(* IEC 61131-3 sources: daoli-st-library/DL_Process (part 9) *)

(* ---- FC_DL_AnodizeBathChargeCalc.st ---- *)
(*
  Component : FC_DL_AnodizeBathChargeCalc
  Category  : DL_Process
  Type      : FC
  Complexity: C2
  VERSION   : v1.0.0
  功能      : 阳极氧化槽法拉第电量核算：Q = I·t，换算电量密度与膜厚，并按电流效率由目标膜厚反算所需时间。
  开源溯源  : 道莅原创 clean-room 自研（无外部代码引用）｜License: MIT
  边界条件  : ① 氧化面积、电流效率、单位电量膜厚系数须 > 1e-9 且效率不超过 100 %，否则返回哨兵 -1；
              ② 电流为 0 时膜厚为 0 且反算时间回 0（合法空工况，xValid 置真）；
              ③ 反算时间不下发负值，目标膜厚 <= 0 时直接回 0。
*)
FUNCTION FC_DL_AnodizeBathChargeCalc : REAL
VAR_INPUT
    fCurrentA     : REAL;   (* 整流器输出电流 [A] Rectifier output current *)
    fAreaDm2      : REAL;   (* 氧化有效面积 [dm²] Effective anodizing area *)
    fTimeS        : REAL;   (* 通电时长 [s] Energizing time *)
    fEffPct       : REAL;   (* 电流效率 [%] Current efficiency *)
    fUmPerAsDm2   : REAL;   (* 单位电量膜厚系数 [μm/(A·s/dm²)] Film thickness per charge density *)
    fThickTargetUm: REAL;   (* 目标膜厚 [μm] Target film thickness *)
END_VAR
VAR_OUTPUT
    fChargeC       : REAL;  (* 累计电量 [C] Accumulated charge *)
    fChgDensAsDm2  : REAL;  (* 电量密度 [A·s/dm²] Charge density *)
    fFilmUm        : REAL;  (* 实测对应膜厚 [μm] Film thickness from charge *)
    fTimeForTargetS: REAL;  (* 达目标膜厚所需时间 [s] Time to reach target thickness *)
    xValid         : BOOL;  (* 计算有效性标志 [-] Calculation valid flag *)
END_VAR
VAR CONSTANT
    DL_EPS      : REAL := 1.0E-9;   (* 除零判定容差 [无量纲] Divide-by-zero tolerance *)
    DL_PCT_BASE : REAL := 100.0;    (* 百分比基准 [%] Percent base *)
    DL_ZERO     : REAL := 0.0;      (* 零常量 [无量纲] Zero constant *)
END_VAR
VAR
    fDensADm2 : REAL;   (* 电流密度 [A/dm²] Current density *)
    fEffUnit  : REAL;   (* 效率折算系数 [-] Efficiency as fraction *)
END_VAR
(* 出口预置：五出口统一预置 *)
fChargeC := 0.0; fChgDensAsDm2 := 0.0; fFilmUm := 0.0; fTimeForTargetS := 0.0; xValid := FALSE;
(* 非有限拦截：自反判 NaN，自身差值判 Inf *)
IF (fCurrentA <> fCurrentA) OR ((fCurrentA - fCurrentA) <> 0.0)
   OR (fAreaDm2 <> fAreaDm2) OR ((fAreaDm2 - fAreaDm2) <> 0.0)
   OR (fTimeS <> fTimeS) OR ((fTimeS - fTimeS) <> 0.0)
   OR (fEffPct <> fEffPct) OR ((fEffPct - fEffPct) <> 0.0)
   OR (fUmPerAsDm2 <> fUmPerAsDm2) OR ((fUmPerAsDm2 - fUmPerAsDm2) <> 0.0) THEN
    FC_DL_AnodizeBathChargeCalc := -1.0;  (* 哨兵 -1：输入非有限 / Sentinel -1 non-finite *)
    RETURN;
END_IF
(* 组态域闸：面积与系数为除子/比例基，电流与时长须非负，效率须在 (0,100] *)
IF (fAreaDm2 <= DL_EPS) OR (fUmPerAsDm2 <= DL_EPS) OR (fEffPct <= DL_ZERO)
   OR (fEffPct > DL_PCT_BASE) OR (fCurrentA < DL_ZERO) OR (fTimeS < DL_ZERO) THEN
    FC_DL_AnodizeBathChargeCalc := -1.0;  (* 哨兵 -1：组态非法 / Sentinel -1 bad config *)
    RETURN;
END_IF
fEffUnit := fEffPct / DL_PCT_BASE;             (* 效率折算 [-] / Efficiency as fraction *)
(* 电量：Q = I·t [C] = [A·s] *)
fChargeC := fCurrentA * fTimeS;
(* 电量密度与电流密度：分母面积已过域闸 *)
fChgDensAsDm2 := fChargeC / fAreaDm2;
fDensADm2 := fCurrentA / fAreaDm2;
(* 膜厚：δ = 电量密度 × 单位膜厚系数 × 电流效率 [μm] *)
fFilmUm := fChgDensAsDm2 * fUmPerAsDm2 * fEffUnit;
(* 反算时间：t = 目标膜厚 / (电流密度 × 系数 × 效率)，电流密度为 0 时回 0 *)
IF (fDensADm2 > DL_EPS) AND (fThickTargetUm > DL_ZERO) THEN
    fTimeForTargetS := fThickTargetUm / (fDensADm2 * fUmPerAsDm2 * fEffUnit);
END_IF
xValid := TRUE;                                (* 链路有效 / Chain valid *)
FC_DL_AnodizeBathChargeCalc := fFilmUm;        (* 返回膜厚 [μm] / Return film thickness *)
END_FUNCTION

(* ---- FC_DL_AnodizeSealBoilTimeCalc.st ---- *)
(*
  Component : FC_DL_AnodizeSealBoilTimeCalc
  Category  : DL_Process
  Type      : FC
  Complexity: C1
  VERSION   : v1.0.0
  功能      : 沸水封孔时间核算：按膜厚乘单位膜厚基准时间，再叠加温度窗口修正，判定 pH/温度窗口与最终封孔合格性。
  开源溯源  : 道莅原创 clean-room 自研（无外部代码引用）｜License: MIT
  边界条件  : ① 膜厚与单位膜厚时间须 > 1e-9，否则返回哨兵 -1；
              ② pH 窗口 5.5~6.5、温度窗口 95~100 °C，任一越窗即判不合格但不拒算；
              ③ 温度修正系数钳位 1.0~2.0，温度偏低延长封孔时间。
*)
FUNCTION FC_DL_AnodizeSealBoilTimeCalc : REAL
VAR_INPUT
    fFilmUm    : REAL;   (* 氧化膜厚 [μm] Oxide film thickness *)
    fBathTempC : REAL;   (* 封孔槽液温度 [°C] Sealing bath temperature *)
    fPh        : REAL;   (* 封孔槽液 pH [-] Sealing bath pH *)
    fMinPerUm  : REAL;   (* 单位膜厚基准封孔时间 [min/μm] Base sealing time per um *)
    fFilmMinUm : REAL;   (* 可封孔最小膜厚 [μm] Minimum sealable film thickness *)
END_VAR
VAR_OUTPUT
    fSealTimeMin : REAL;  (* 封孔时间 [min] Sealing time *)
    fTempCoef    : REAL;  (* 温度修正系数 [-] Temperature correction coefficient *)
    xWindowOk    : BOOL;  (* pH 与温度窗口合格标志 [-] Window valid flag *)
    xQualified   : BOOL;  (* 封孔合格标志 [-] Sealing qualified flag *)
    xValid       : BOOL;  (* 计算有效性标志 [-] Calculation valid flag *)
END_VAR
VAR CONSTANT
    DL_EPS      : REAL := 1.0E-9;   (* 除零判定容差 [无量纲] Divide-by-zero tolerance *)
    DL_PH_LO    : REAL := 5.5;      (* pH 窗口下限 [-] pH window lower bound *)
    DL_PH_HI    : REAL := 6.5;      (* pH 窗口上限 [-] pH window upper bound *)
    DL_TMP_LO   : REAL := 95.0;     (* 温度窗口下限 [°C] Temperature window lower bound *)
    DL_TMP_HI   : REAL := 100.0;    (* 温度窗口上限 [°C] Temperature window upper bound *)
    DL_TMP_REF  : REAL := 100.0;    (* 温度修正基准 [°C] Temperature reference *)
    DL_TMP_SLOPE: REAL := 0.25;     (* 每 10 °C 温度修正量 [-] Slope per 10 degC *)
    DL_COEF_MAX : REAL := 2.0;      (* 温度修正上限 [-] Temperature coefficient clamp *)
END_VAR
VAR
    fGapC : REAL;   (* 相对基准温度的温差 [°C] Temperature gap from reference *)
END_VAR
(* 出口预置：五出口统一预置 *)
fSealTimeMin := 0.0; fTempCoef := 1.0; xWindowOk := FALSE; xQualified := FALSE; xValid := FALSE;
(* 非有限拦截：自反判 NaN，自身差值判 Inf *)
IF (fFilmUm <> fFilmUm) OR ((fFilmUm - fFilmUm) <> 0.0)
   OR (fBathTempC <> fBathTempC) OR ((fBathTempC - fBathTempC) <> 0.0)
   OR (fPh <> fPh) OR ((fPh - fPh) <> 0.0) THEN
    FC_DL_AnodizeSealBoilTimeCalc := -1.0;  (* 哨兵 -1：输入非有限 / Sentinel -1 non-finite *)
    RETURN;
END_IF
(* 组态域闸：膜厚与单位膜厚时间均为比例基 *)
IF (fFilmUm < DL_EPS) OR (fMinPerUm <= DL_EPS) THEN
    FC_DL_AnodizeSealBoilTimeCalc := -1.0;  (* 哨兵 -1：组态非法 / Sentinel -1 bad config *)
    RETURN;
END_IF
(* 窗口判定：pH 与温度双窗口，任一越窗即判不合格（不拒算，便于上位诊断） *)
IF (fPh >= DL_PH_LO) AND (fPh <= DL_PH_HI)
   AND (fBathTempC >= DL_TMP_LO) AND (fBathTempC <= DL_TMP_HI) THEN
    xWindowOk := TRUE;
END_IF
(* 温度修正：低于基准温度每 10 °C 延长 25 %，双侧钳位 *)
fGapC := DL_TMP_REF - fBathTempC;
IF fGapC > 0.0 THEN
    fTempCoef := 1.0 + (fGapC / 10.0) * DL_TMP_SLOPE;
ELSE
    fTempCoef := 1.0;                       (* 达到或高于基准：不缩短，防欠封 *)
END_IF
IF fTempCoef > DL_COEF_MAX THEN
    fTempCoef := DL_COEF_MAX;               (* 上限钳位 [-] / Upper clamp *)
END_IF
(* 封孔时间：t = 膜厚 × 单位膜厚时间 × 温度修正，分母均已过域闸 *)
fSealTimeMin := fFilmUm * fMinPerUm * fTempCoef;
(* 合格判定：窗口合格且膜厚达可封孔最小值 *)
xQualified := xWindowOk AND (fFilmUm >= fFilmMinUm);
xValid := TRUE;                             (* 链路有效 / Chain valid *)
FC_DL_AnodizeSealBoilTimeCalc := fSealTimeMin;  (* 返回封孔时间 [min] / Return sealing minutes *)
END_FUNCTION

(* ---- FC_DL_AustenitizeHoldTimeCalc.st ---- *)
(*
  Component : FC_DL_AustenitizeHoldTimeCalc
  Category  : DL_Process
  Type      : FC
  Complexity: C2
  VERSION   : v1.0.0
  功能      : 奥氏体化保温时间核算：按有效厚度乘以单位厚度基准时间，再叠加厚度分段系数、升温速率修正与目标温度修正。
  开源溯源  : 道莅原创 clean-room 自研（无外部代码引用）｜License: MIT
  边界条件  : ① 有效厚度/升温速率/单位厚度时间均须 > 1e-9，否则返回哨兵 -1；
              ② 厚度分三段（<=25 / <=50 / >50 mm），系数逐段离散，段内不插值；
              ③ 升温速率修正与温度修正均双侧钳位，防经验式外推发散。
*)
FUNCTION FC_DL_AustenitizeHoldTimeCalc : REAL
VAR_INPUT
    fThkMm      : REAL;   (* 工件有效厚度 [mm] Effective thickness *)
    fRateCmin   : REAL;   (* 实际升温速率 [°C/min] Actual heating rate *)
    fRateRefCmin: REAL;   (* 参考升温速率（分段基准） [°C/min] Reference heating rate *)
    fTargetC    : REAL;   (* 目标奥氏体化温度 [°C] Target austenitizing temperature *)
    fTempRefC   : REAL;   (* 参考目标温度（分段基准） [°C] Reference target temperature *)
    fMinPerMm   : REAL;   (* 单位厚度基准保温时间 [min/mm] Base hold time per mm *)
END_VAR
VAR_OUTPUT
    fHoldMin   : REAL;    (* 保温时间计算结果 [min] Computed hold time *)
    fThkCoef   : REAL;    (* 厚度分段系数 [-] Thickness segment coefficient *)
    fRateCoef  : REAL;    (* 升温速率修正系数 [-] Heating rate correction coefficient *)
    xValid     : BOOL;    (* 计算有效性标志 [-] Calculation valid flag *)
END_VAR
VAR CONSTANT
    DL_EPS       : REAL := 1.0E-9;   (* 除零判定容差 [无量纲] Divide-by-zero tolerance *)
    DL_RATE_MIN  : REAL := 0.80;     (* 速率修正下限 [-] Rate correction lower clamp *)
    DL_RATE_MAX  : REAL := 1.30;     (* 速率修正上限 [-] Rate correction upper clamp *)
    DL_TEMP_K    : REAL := 0.002;    (* 目标温度每 °C 修正斜率 [1/°C] Temperature slope *)
    DL_THK_MID   : REAL := 25.0;     (* 厚度分段第一界 [mm] First thickness boundary *)
    DL_THK_HIGH  : REAL := 50.0;     (* 厚度分段第二界 [mm] Second thickness boundary *)
END_VAR
(* 出口预置：全出口统一预置 *)
fHoldMin := 0.0; fThkCoef := 1.0; fRateCoef := 1.0; xValid := FALSE;
(* 非有限拦截：自反判 NaN，自身差值判 Inf *)
IF (fThkMm <> fThkMm) OR ((fThkMm - fThkMm) <> 0.0)
   OR (fRateCmin <> fRateCmin) OR ((fRateCmin - fRateCmin) <> 0.0)
   OR (fRateRefCmin <> fRateRefCmin) OR ((fRateRefCmin - fRateRefCmin) <> 0.0)
   OR (fTargetC <> fTargetC) OR ((fTargetC - fTargetC) <> 0.0)
   OR (fTempRefC <> fTempRefC) OR ((fTempRefC - fTempRefC) <> 0.0)
   OR (fMinPerMm <> fMinPerMm) OR ((fMinPerMm - fMinPerMm) <> 0.0) THEN
    FC_DL_AustenitizeHoldTimeCalc := -1.0;  (* 哨兵 -1：输入非有限 / Sentinel -1 non-finite *)
    RETURN;
END_IF
(* 组态域闸：厚度、实际升温速率、单位厚度时间三者为除子或比例基 *)
IF (fThkMm <= DL_EPS) OR (fRateCmin <= DL_EPS) OR (fMinPerMm <= DL_EPS) THEN
    FC_DL_AustenitizeHoldTimeCalc := -1.0;  (* 哨兵 -1：组态非法 / Sentinel -1 bad config *)
    RETURN;
END_IF
(* 厚度分段系数：三段离散，段内不插值，防止经验式在厚壁区外推 *)
IF fThkMm <= DL_THK_MID THEN
    fThkCoef := 1.00;                       (* 薄件段 [-] / Thin section *)
ELSIF fThkMm <= DL_THK_HIGH THEN
    fThkCoef := 1.15;                       (* 中厚段 [-] / Medium section *)
ELSE
    fThkCoef := 1.35;                       (* 厚壁段（心部透热滞后） [-] / Thick section *)
END_IF
(* 升温速率修正：升温越慢，组织转变越充分，保温时间可缩短，双侧钳位 *)
fRateCoef := fRateRefCmin / fRateCmin;
IF fRateCoef < DL_RATE_MIN THEN
    fRateCoef := DL_RATE_MIN;               (* 下限钳位 [-] / Lower clamp *)
ELSIF fRateCoef > DL_RATE_MAX THEN
    fRateCoef := DL_RATE_MAX;               (* 上限钳位 [-] / Upper clamp *)
END_IF
(* 目标温度修正：温度偏低需延长保温 *)
IF fTargetC > fTempRefC THEN
    fHoldMin := fMinPerMm * fThkMm * fThkCoef * fRateCoef;
    fHoldMin := fHoldMin * (1.0 - (fTargetC - fTempRefC) * DL_TEMP_K);
ELSE
    fHoldMin := fMinPerMm * fThkMm * fThkCoef * fRateCoef;
    fHoldMin := fHoldMin * (1.0 + (fTempRefC - fTargetC) * DL_TEMP_K);
END_IF
(* 结果下钳位：保温时间不得为负，防温度修正项越界 *)
IF fHoldMin < DL_EPS THEN
    fHoldMin := DL_EPS;                     (* 非负钳位 [min] / Non-negative clamp *)
END_IF
xValid := TRUE;                             (* 链路有效 / Chain valid *)
FC_DL_AustenitizeHoldTimeCalc := fHoldMin;  (* 返回保温时间 [min] / Return hold minutes *)
END_FUNCTION

(* ---- FC_DL_BallMillPowerDrawCalc.st ---- *)
(*
  Name: FC_DL_BallMillPowerDrawCalc
  Category: DL_Process
  Version: 1.0.0
  Round: R89 / 2026-11-25
  开源溯源：clean-room 自研（族 矿山破碎筛分，ST 开源生态实测 0 命中，无外部代码引入）
  功能：球磨机轴功率与比能耗估算（筒径/筒长/转速率/装球率经验幂律），并折算单位给矿能耗。
  边界条件：① 五入参全部过非有限闸，任一非有限返回哨兵 -1；
            ② 筒径 0.5~8 m、筒长 0.5~15 m、临界转速率 30~100 %、装球率 10~55 % 为工程域，越域返回哨兵 -1；
            ③ 给矿量为 0 属正常运行工况（空转），比能耗输出 0 而不判非法，功率照常有效；
            ④ 幂次 2.5 以 D·D·SQRT(D) 展开实现，不引入 EXPT 原语（R140 委托纪律）。
  量纲自证：K[kW/m^3.5] × D^2.5[m^2.5] × L[m] = kW；转速率与装球率为无量纲百分比折算。
*)
FUNCTION FC_DL_BallMillPowerDrawCalc : REAL
VAR_INPUT
    fMillDiaM : REAL;        (* 磨机筒体有效内径 [m] Mill effective diameter [m] *)
    fMillLenM : REAL;        (* 磨机筒体有效长度 [m] Mill effective length [m] *)
    fSpeedPct : REAL;        (* 临界转速百分比 [%] Percent of critical speed [%] *)
    fMediaLoadPct : REAL;    (* 装球率（磨机容积占比） [%] Ball charge volume ratio [%] *)
    fFeedTph : REAL;         (* 给矿量 [t/h] Feed rate [t/h] *)
END_VAR
VAR_OUTPUT
    fPowerKW : REAL;         (* 磨机轴功率 [kW] Mill shaft power [kW] *)
    fSpecificKWhT : REAL;    (* 单位给矿能耗 [kWh/t] Specific energy per tonne [kWh/t] *)
    xValid : BOOL;           (* 计算有效性标志 [-] Calculation valid flag *)
END_VAR
VAR CONSTANT
    DL_EPS : REAL := 1.0E-9;        (* 除零判定容差 [-] Divide-by-zero tolerance *)
    DL_K_POWER : REAL := 26.0;      (* 功率经验系数 [kW/m^3.5] Empirical power coefficient *)
    DL_D_MIN : REAL := 0.5;         (* 筒径下限 [m] Diameter floor [m] *)
    DL_D_MAX : REAL := 8.0;         (* 筒径上限 [m] Diameter ceiling [m] *)
    DL_L_MIN : REAL := 0.5;         (* 筒长下限 [m] Length floor [m] *)
    DL_L_MAX : REAL := 15.0;        (* 筒长上限 [m] Length ceiling [m] *)
    DL_SPD_MIN : REAL := 30.0;      (* 转速率下限 [%] Speed ratio floor [%] *)
    DL_SPD_MAX : REAL := 100.0;     (* 转速率上限 [%] Speed ratio ceiling [%] *)
    DL_MED_MIN : REAL := 10.0;      (* 装球率下限 [%] Media load floor [%] *)
    DL_MED_MAX : REAL := 55.0;      (* 装球率上限 [%] Media load ceiling [%] *)
    DL_PCT : REAL := 100.0;         (* 百分数基准 [%] Percent base *)
END_VAR
VAR
    fD25 : REAL;    (* 筒径 2.5 次幂 [m^2.5] Diameter to the power 2.5 *)
    fKspd : REAL;   (* 转速率折算系数 [-] Speed ratio factor *)
    fKmed : REAL;   (* 装球率折算系数 [-] Media load factor *)
END_VAR
(* 出口预置：三出口统一预置（R256） *)
fPowerKW := 0.0; fSpecificKWhT := 0.0; xValid := FALSE;
(* 非有限闸：NaN 自反判 + Inf 差值自减判，五入参全枚举 *)
IF (fMillDiaM <> fMillDiaM) OR ((fMillDiaM - fMillDiaM) <> 0.0)
   OR (fMillLenM <> fMillLenM) OR ((fMillLenM - fMillLenM) <> 0.0)
   OR (fSpeedPct <> fSpeedPct) OR ((fSpeedPct - fSpeedPct) <> 0.0)
   OR (fMediaLoadPct <> fMediaLoadPct) OR ((fMediaLoadPct - fMediaLoadPct) <> 0.0)
   OR (fFeedTph <> fFeedTph) OR ((fFeedTph - fFeedTph) <> 0.0) THEN
    FC_DL_BallMillPowerDrawCalc := -1.0;    (* 哨兵 -1：入参非有限 / Sentinel -1, non-finite input *)
    RETURN;
END_IF
(* 组态域闸：几何与工艺参数逐项定域，给矿量允许为 0（空转） *)
IF (fMillDiaM < DL_D_MIN) OR (fMillDiaM > DL_D_MAX)
   OR (fMillLenM < DL_L_MIN) OR (fMillLenM > DL_L_MAX)
   OR (fSpeedPct < DL_SPD_MIN) OR (fSpeedPct > DL_SPD_MAX)
   OR (fMediaLoadPct < DL_MED_MIN) OR (fMediaLoadPct > DL_MED_MAX)
   OR (fFeedTph < 0.0) THEN
    FC_DL_BallMillPowerDrawCalc := -1.0;    (* 哨兵 -1：组态非法 / Sentinel -1, bad configuration *)
    RETURN;
END_IF
(* 幂次展开：D^2.5 = D·D·√D，量纲 m^2.5 *)
fD25 := fMillDiaM * fMillDiaM * SQRT(fMillDiaM);
(* 两百分比折算为无量纲系数 *)
fKspd := fSpeedPct / DL_PCT;
fKmed := fMediaLoadPct / DL_PCT;
(* 轴功率：K[kW/m^3.5] × D^2.5 × L × kspd × kmed，量纲收敛为 kW *)
fPowerKW := DL_K_POWER * fD25 * fMillLenM * fKspd * fKmed;
(* 比能耗：给矿为 0 时输出 0（除零保护，且空转不产比能耗事实） *)
IF fFeedTph > DL_EPS THEN
    fSpecificKWhT := fPowerKW / fFeedTph;   (* kW ÷ (t/h) = kWh/t *)
ELSE
    fSpecificKWhT := 0.0;                   (* 空转：无比能耗 / No specific energy at no feed *)
END_IF
xValid := TRUE;                             (* 链路有效 / Chain valid *)
FC_DL_BallMillPowerDrawCalc := fPowerKW;
END_FUNCTION

(* ---- FC_DL_BeamToppleRiskChk.st ---- *)
(*
  ============================================================
  组件名 : FC_DL_BeamToppleRiskChk
  分类   : DL_Process
  功能   : 横梁倾覆风险校核，按重心偏心放大力矩后折算横梁承载利用率并给出风险位
  复杂度 : C1
  版本   : 1.0.1
  作者   : 道莅工业代码库工厂 / R81
  日期   : 2026-11-24
  开源溯源 : clean-room（no upstream）—— 依据公开工程公式自研，未复制任何上游实现
  红线自检 : R1 无GVL/R2 无物理地址/R3 纯IEC/R4 防除零/R5 双语注释
  接口说明 :
      偏心系数 = 1 + |重心偏移|/横梁深度（v1.0.1 取绝对值：负偏移同样放大倾覆风险，
      修正原带符号实现导致负偏移时利用率被低估、风险漏报的缺陷），偏心为零时系数为 1。
      |重心偏移| > 梁深/2 视为不可信组态，直接置 bValid=FALSE 返回。
      有效载荷 = 载荷 * 偏心系数；利用率超过 85% 即判倾覆风险。
      利用率不做 100% 上限截断，超过 100% 的信息对诊断有价值，由调用侧自行显示。
  ============================================================
*)
FUNCTION FC_DL_BeamToppleRiskChk : BOOL
VAR_INPUT
    bEnable      : BOOL; // 使能：TRUE 时校核 / Enable: TRUE to check
    bErr         : BOOL; // 外部故障：TRUE 时立即退出并置结果无效 / External fault: TRUE aborts with invalid result
    rLoadKg      : REAL; // 实际载荷质量 [kg] / actual load mass [kg]
    rBeamCapKg   : REAL; // 横梁额定承载质量 [kg] / rated load capacity of the beam [kg]
    rCgOffset_mm : REAL; // 载荷重心相对横梁中心的偏移 [mm] / load centre of gravity offset from the beam centre [mm]
    rBeamDepth_mm : REAL; // 横梁截面深度 [mm] / beam section depth [mm]
END_VAR
VAR_OUTPUT
    rEccFactor : REAL; // 偏心放大系数 [无量纲] / eccentricity amplification factor [dimensionless]
    rEffLoadKg : REAL; // 折算有效载荷质量 [kg] / equivalent effective load mass [kg]
    rUtilPct   : REAL; // 承载利用率 [%] / utilisation of the rated capacity [percent]
    bRisk      : BOOL; // 倾覆风险：TRUE 表示利用率超过门限 / topple risk, TRUE when utilisation exceeds the limit
    bValid     : BOOL; // 输出有效：TRUE 表示结果可用 / Output valid
END_VAR
VAR CONSTANT
    DL_R_MAX    : REAL := 3.0E38; // 实数上界，用于拦截 Inf [无量纲] / real upper bound used to reject infinity [dimensionless]
    DL_EPS      : REAL := 1.0E-12; // 除零判定阈值 [无量纲] / division guard threshold [dimensionless]
    DL_RISK_PCT : REAL := 85.0;   // 倾覆风险门限 [%] / topple risk threshold [percent]
    DL_PCT      : REAL := 100.0;  // 百分数换算系数 [无量纲] / percentage scaling factor [dimensionless]
END_VAR
VAR
    _bFin : BOOL := FALSE; // 输入有限性判定结果 / input finiteness verdict
END_VAR

    // 段 1｜出口预置
    rEccFactor := 1.0;
    rEffLoadKg := 0.0;
    rUtilPct := 0.0;
    bRisk := FALSE;
    bValid := FALSE;
    // 段 2｜使能闸与外部故障闸
    IF NOT bEnable THEN
        RETURN;
    END_IF;
    IF bErr THEN
        RETURN;
    END_IF;
    // 段 3｜非有限闸
    _bFin := (rLoadKg = rLoadKg) AND (ABS(rLoadKg) <= DL_R_MAX) AND (rBeamCapKg = rBeamCapKg) AND (ABS(rBeamCapKg) <= DL_R_MAX) AND (rCgOffset_mm = rCgOffset_mm) AND (ABS(rCgOffset_mm) <= DL_R_MAX) AND (rBeamDepth_mm = rBeamDepth_mm) AND (ABS(rBeamDepth_mm) <= DL_R_MAX);
    IF NOT _bFin THEN
        RETURN;
    END_IF;
    // 段 4｜域闸：承载与横梁深度必须为正，载荷不得为负
    IF (ABS(rBeamCapKg) <= DL_EPS) OR (ABS(rBeamDepth_mm) <= DL_EPS) THEN
        RETURN;
    END_IF;
    IF (rBeamCapKg < 0.0) OR (rLoadKg < 0.0) OR (rBeamDepth_mm < 0.0) THEN
        RETURN;
    END_IF;
    // 段 4b｜偏心量域闸：|偏移| 超过梁深一半即视为不可信组态，直接置无效退出（R81 闸席 FAIL(LOGIC) 修法）
    IF ABS(rCgOffset_mm) > (rBeamDepth_mm * 0.5) THEN
        RETURN;
    END_IF;
    // 段 5｜偏心放大系数：取偏移绝对值，负偏移（重心偏向另一侧）同样放大倾覆风险 / use absolute offset
    rEccFactor := 1.0 + ABS(rCgOffset_mm) / rBeamDepth_mm;
    // 段 6｜有效载荷与利用率
    rEffLoadKg := rLoadKg * rEccFactor;
    rUtilPct := rEffLoadKg / rBeamCapKg * DL_PCT;
    // 段 7｜风险位：严格大于门限才置位，等于门限视为可控
    IF rUtilPct > DL_RISK_PCT THEN
        bRisk := TRUE;
    ELSE
        bRisk := FALSE;
    END_IF;
    bValid := TRUE;
    FC_DL_BeamToppleRiskChk := bValid;
END_FUNCTION

(* ---- FC_DL_BeamWarpLengthCalc.st ---- *)
(*
  DL Factory R83 | FC_DL_BeamWarpLengthCalc
  功能：按边盘与轴芯直径、纱线直径算经轴卷绕层数、可卷经纱长度与总根数。
  开源溯源：无（clean-room 自研，依据公开工艺公式，来源=行业通用公式，许可证=MIT，借鉴点=公式结构）
  规则：R1-R21 全遵守
*)
FUNCTION FC_DL_BeamWarpLengthCalc : REAL
VAR_INPUT
    fFlangeDiaMm : REAL; // 经轴边盘直径 [mm] / Beam flange diameter [mm]
    fBarrelDiaMm : REAL; // 经轴轴芯直径 [mm] / Beam barrel diameter [mm]
    fYarnDiaMm   : REAL; // 单根经纱直径（即单层卷绕厚度）[mm] / Yarn diameter, layer thickness [mm]
    fWarpDensity : REAL; // 经密（每 cm 根数）[根/cm] / Warp density [ends/cm]
    fBeamWidthMm : REAL; // 经轴卷绕幅宽 [mm] / Beam winding width [mm]
END_VAR
VAR_OUTPUT
    fLengthM : REAL; // 可卷绕经纱总长 [m] / Windable warp length [m]
    iLayers  : INT;  // 可卷绕层数 [层] / Number of wound layers [-]
    diEnds   : DINT; // 经纱总根数 [根] / Total warp ends [-]
    xValid   : BOOL; // 计算有效性标志 / Calculation validity flag
END_VAR
VAR
    fOuterMm : REAL; // 满轴外径 [mm] / Fully wound outer diameter [mm]
    fAvgMm   : REAL; // 平均卷绕直径 [mm] / Mean winding diameter [mm]
    fRadialMm: REAL; // 径向可卷厚度 [mm] / Available radial thickness [mm]
END_VAR
// 出口预置：四出口统一预置（R256）
fLengthM := 0.0; iLayers := 0; diEnds := 0; xValid := FALSE;
// 非有限拦截 + 量纲次序 + 分母零闸（R4/R20/R21）
IF NOT (fFlangeDiaMm > -1.0E30 AND fFlangeDiaMm < 1.0E30) OR NOT (fBarrelDiaMm > -1.0E30 AND fBarrelDiaMm < 1.0E30) OR NOT (fYarnDiaMm > -1.0E30 AND fYarnDiaMm < 1.0E30) OR NOT (fWarpDensity > -1.0E30 AND fWarpDensity < 1.0E30) OR NOT (fBeamWidthMm > -1.0E30 AND fBeamWidthMm < 1.0E30) OR fFlangeDiaMm <= fBarrelDiaMm OR ABS(fYarnDiaMm) <= 1.0E-9 OR fWarpDensity <= 0.0 OR fBeamWidthMm <= 0.0 THEN
    FC_DL_BeamWarpLengthCalc := -1.0; RETURN;   // 哨兵 -1：非有限或量纲/直径次序越界 / Sentinel -1
END_IF
// 径向可卷厚度：(边盘 - 轴芯) ÷ 2，单边径向空间 [mm]
fRadialMm := (fFlangeDiaMm - fBarrelDiaMm) / 2.0;   // 径向厚度 [mm] / Radial thickness [mm]
// 层数：向下取整（禁 TRUNC+1 向上取整写法，R28）
iLayers := REAL_TO_INT(fRadialMm / fYarnDiaMm);     // 满层数 [层] / Full layers [-]
// 平均卷绕直径：轴芯与满轴外径的中径，外径 = 轴芯 + 层数 × 纱径（mm）
fOuterMm := fBarrelDiaMm + INT_TO_REAL(iLayers) * fYarnDiaMm; // 满轴外径 [mm] / Outer diameter [mm]
fAvgMm   := (fBarrelDiaMm + fOuterMm) / 2.0;                  // 平均直径 [mm] / Mean diameter [mm]
// 纱长：层数 × π × 平均直径，mm ÷ 1000 得 m（量纲自洽）
IF iLayers > 0 THEN
    fLengthM := 3.14159265358979 * fAvgMm * INT_TO_REAL(iLayers) / 1000.0; // 卷绕长度 [m]
ELSE
    fLengthM := 0.0;                // 不足一层不可卷绕 / Not even one layer, zero length
END_IF
// 经纱根数：根/cm × 幅宽(cm) = 根；幅宽 mm ÷ 10 = cm（量纲自洽）
diEnds := REAL_TO_DINT(fWarpDensity * fBeamWidthMm / 10.0); // 总根数 [根] / Total ends [-]
xValid := TRUE;                                             // 链路有效 / Chain valid
FC_DL_BeamWarpLengthCalc := fLengthM;                       // 返回可卷长度 [m] / Return length [m]
END_FUNCTION

(* ---- FC_DL_BeerCoolingLoadCalc.st ---- *)
// FC_DL_BeerCoolingLoadCalc v1.0.0
// 开源溯源：clean-room 自研（族 DL_Process，ST 生态实测 0 命中，无外部代码引入）
(*
  功能: 冷却负荷：体积流量 = 流量[hL/h]·100/1000 [m³/h]，质量流量 = 体积流量·ρ/3600 [kg/s]，
        显热负荷 = 质量流量·cp·(进料 − 出料) [kW]（kJ/s = kW），总冷负荷 = 显热 + 发酵放热。
  邻件/码位: 与 FC_DL_DiacetylRestWindowCalc、FC_DL_KegFillingCounterPressureCalc 同属后段冷工链；
             16#0002_9239 = 非有限、流量/密度/比热非正、出料不低于进料或发酵热为负拒收。
*)
FUNCTION FC_DL_BeerCoolingLoadCalc : REAL
VAR_INPUT
    fFlow        : REAL := 200.0;   // 流量 [hL/h]，域 > 0 / Flow rate [hL/h]
    fTempIn      : REAL := 12.0;    // 进料温度 [°C] / Inlet temperature [degC]
    fTempOut     : REAL := 2.0;     // 出料温度 [°C]，域 < 进料 / Outlet temperature [degC]
    fCp          : REAL := 3.85;    // 比热 [kJ/(kg·K)]，域 > 0 / Specific heat [kJ/(kg K)]
    fDensity     : REAL := 1010.0;  // 密度 [kg/m³]，域 > 0 / Density [kg/m^3]
    fFermentHeat : REAL := 5.0;     // 发酵放热 [kW]，域 >= 0 / Fermentation heat [kW]
END_VAR
VAR_OUTPUT
    fCoolLoad : REAL;               // 总冷负荷 [kW] / Total cooling load [kW]
    bValid    : BOOL;               // 结果有效回执 [-] / Result validity receipt
    uErrorId  : UDINT;              // 事件码，0 = 无事件 / Event code
END_VAR
VAR
    fMassFlow : REAL := 0.0;        // 质量流量 [kg/s] / Mass flow [kg/s]
END_VAR
// 段 0：全路径出口安全缺省 / Safe defaults on all outlets
fCoolLoad := 0.0;                   // 冷负荷缺省零 / Cooling load default zero
bValid := FALSE;                    // 有效回执预清 / Validity preset clear
uErrorId := 16#0000;                // 事件码预清 / Event code preset clear
FC_DL_BeerCoolingLoadCalc := 0.0;   // 返回值缺省零（镜像冷负荷）/ Return default zero
// 段 1：非有限闸（六入参全枚举）/ Non-finite gate over all inputs
IF (fFlow <> fFlow) OR (fTempIn <> fTempIn) OR (fTempOut <> fTempOut)
   OR (fCp <> fCp) OR (fDensity <> fDensity) OR (fFermentHeat <> fFermentHeat)
   OR (ABS(fFlow) >= 3.0E38) OR (ABS(fTempIn) >= 3.0E38) OR (ABS(fTempOut) >= 3.0E38)
   OR (ABS(fCp) >= 3.0E38) OR (ABS(fDensity) >= 3.0E38) OR (ABS(fFermentHeat) >= 3.0E38) THEN
    uErrorId := 16#0002_9239;   // 入参非有限拒收 / Non-finite input reject
    RETURN;
END_IF
// 段 2：域闸（流量/密度/比热为正 + 出料低于进料 + 发酵热非负，R4）/ Domain gate
IF (fFlow <= 1.0E-6) OR (fDensity <= 1.0E-6) OR (fCp <= 1.0E-6) THEN
    uErrorId := 16#0002_9239;   // 流量、密度或比热非正 / Non-positive flow, density or capacity
    RETURN;
END_IF
IF fTempOut >= fTempIn THEN
    uErrorId := 16#0002_9239;   // 出料不低于进料，无冷却需求 / Outlet not colder than inlet
    RETURN;
END_IF
IF fFermentHeat < 0.0 THEN
    uErrorId := 16#0002_9239;   // 发酵放热为负 / Negative fermentation heat
    RETURN;
END_IF
// 段 3：主计算（体积→质量流量 → 显热 → 总负荷）/ Main computation
fMassFlow := fFlow * 100.0 / 1000.0 * fDensity / 3600.0;        // 质量流量 [kg/s] / Mass flow
fCoolLoad := fMassFlow * fCp * (fTempIn - fTempOut) + fFermentHeat;     // 总冷负荷 [kW] / Total load
// 段 4：出口闸（非有限复核 + 正数复核）/ Outlet gate
IF (fCoolLoad <> fCoolLoad) OR (ABS(fCoolLoad) >= 3.0E38) OR (fCoolLoad <= 0.0) THEN
    fCoolLoad := 0.0;           // 复核失败回缺省 / Fallback on recheck failure
    uErrorId := 16#0002_9239;   // 出口复核拒收 / Output recheck reject
    RETURN;
END_IF
bValid := TRUE;                 // 有效回执 / Validity receipt
FC_DL_BeerCoolingLoadCalc := fCoolLoad;         // 返回值镜像总冷负荷 / Return mirrors load
END_FUNCTION

(* ---- FC_DL_BeltPressLoadRate.st ---- *)
(*
  道莅工业代码库 / Daoli Industrial ST Library
  组件: FC_DL_BeltPressLoadRate
  分类: DL_Process
  开源溯源: 无（clean-room 工程公式自研；参考公开工艺计算公式，未复制任何受版权保护代码）
  许可证: 本项目自有 (MIT)
  功能: 带式压滤机单位滤带面积固体比负荷计算与过载判定
*)
FUNCTION FC_DL_BeltPressLoadRate : BOOL
VAR_INPUT
    rDsKgH : REAL; // 干固体处理量 [kg/h] / dry solids throughput
    rBeltWidthM : REAL; // 滤带有效宽度 [m] / effective belt width
    rBeltSpeedMmin : REAL; // 滤带线速度 [m/min] / belt linear speed
END_VAR
VAR_OUTPUT
    rLoadKgM2h : REAL; // 比负荷 [kg/(m2·h)] / specific solids loading
    bValid : BOOL; // 结果有效位 [-] / result valid flag
    bOver : BOOL; // 过载标志（>500 kg/(m2·h)）[-] / overload flag
    iErrCode : INT; // 事件码 0=正常 1=滤带面积非法 2=结果非有限 / event code
END_VAR
VAR CONSTANT
    rMinPerHour : REAL := 60.0; // 每小时分钟数 [min/h] / minutes per hour
    rLoadHi : REAL := 500.0; // 比负荷过载门槛 [kg/(m2·h)] / overload threshold
END_VAR
VAR
    rAreaM2h : REAL; // 滤带处理面积速率 [m2/h] / belt area rate
    rLoadRaw : REAL; // 未限幅比负荷 [kg/(m2·h)] / unlimited specific loading
END_VAR

    // —— 段 0：全路径预清 —— //
    rAreaM2h := 0.0;
    rLoadRaw := 0.0;
    rLoadKgM2h := 0.0;
    bValid := FALSE;
    bOver := FALSE;
    iErrCode := 0;
    FC_DL_BeltPressLoadRate := FALSE;
    // —— 段 1：分母闸（滤带面积速率 = 宽 × 速 × 60） —— //
    rAreaM2h := rBeltWidthM * rBeltSpeedMmin * rMinPerHour; // 面积速率 [m2/h] / belt area rate
    IF (rBeltWidthM <= 0.0) OR (rAreaM2h <= 0.0) THEN
        iErrCode := 1; // 滤带面积速率非法，比负荷无定义 / invalid belt area rate
        RETURN;
    END_IF;
    // —— 段 2：量纲链 (kg/h)/(m2/h) = kg/(m2·h) —— //
    rLoadRaw := rDsKgH / rAreaM2h; // 比负荷 [kg/(m2·h)] / specific loading
    IF ABS(rLoadRaw) > 1.0E15 THEN
        iErrCode := 2; // 结果非有限，强制归零 / non-finite result, forced to zero
        RETURN;
    END_IF;
    // —— 段 3：负值防御与过载判定 —— //
    IF rLoadRaw < 0.0 THEN
        rLoadKgM2h := 0.0; // 负干固体防御 / negative dry solids guard
    ELSE
        rLoadKgM2h := rLoadRaw;
    END_IF;
    bOver := rLoadKgM2h > rLoadHi; // 过载判定 [-] / overload test
    bValid := TRUE;
    FC_DL_BeltPressLoadRate := TRUE;
END_FUNCTION

(* ---- FC_DL_BentoniteAdditiveCalc.st ---- *)
(*
 * FC_DL_BentoniteAdditiveCalc | C2 | DL_Process
 * 功能：按亚甲基蓝吸附量差额计算膨润土补加比例与补加量       单位：吸附量 [mL/100g]、比例 [%]、流量 [kg/h]、效率 [%]
 * 工况边界：经验系数 0.15 %/(mL/100g)（spec 采纳值），仅适用于湿型砂单一膨润土体系；实测值已达或超过目标时补加量为 0（xNeedAdd=FALSE，不判故障）；砂处理量须 ≥0、效率须在 (0,100] %
 * 代数值回代：mb=35、target=40 → deficit=5；addPct=5×0.15=0.75 %；sandRate=120000 kg/h → 补加 900 kg/h（spec 采纳 0.15 系数回代值 900 kg/h，一致）
 * 系数修正说明：spec 初版给 addKgH = sandRate×(deficit/100)×(100/eff)，回代得 9231 kg/h 明显超出工艺量级，spec 已明确改用 0.15 系数，本件按采纳值实现
 * 开源溯源：clean-room 自研，未复制任何第三方代码（无外部来源）
 *)
FUNCTION FC_DL_BentoniteAdditiveCalc : BOOL
VAR_INPUT
    rMbValueMl    : REAL := 35.0;      // 实测亚甲基蓝吸附量 | measured methylene blue adsorption [mL/100g]
    rMbTarget     : REAL := 40.0;      // 目标亚甲基蓝吸附量 | target methylene blue adsorption [mL/100g]
    rSandRateKgH  : REAL := 120000.0;  // 砂处理量 | sand throughput [kg/h]
    rEffPct       : REAL := 65.0;      // 膨润土有效利用率 | bentonite effective utilisation [%]
END_VAR
VAR_OUTPUT
    rDeficitMb    : REAL;              // 吸附量差额（目标−实测）| adsorption deficit, target minus measured [mL/100g]
    rAddPct       : REAL;              // 补加比例 | additive ratio [%]
    rBentoniteKgH : REAL;              // 膨润土补加量 | bentonite additive rate [kg/h]
    xNeedAdd      : BOOL;              // 需要补加（差额 >0）| additive required, deficit above zero
    xValid        : BOOL;              // 输出有效 | outputs valid
    nFaultCode    : INT;               // 0=无 / 9713=输入非法 | 0 none, 9713 illegal input
END_VAR
VAR
    xFinMb   : BOOL;                   // 实测值有限性 | measured value is finite
    xFinTg   : BOOL;                   // 目标值有限性 | target is finite
    xFinRate : BOOL;                   // 处理量有限性 | throughput is finite
    xFinEff  : BOOL;                   // 效率有限性 | efficiency is finite
END_VAR
VAR CONSTANT
    DL_BAC_PCT_PER_ML : REAL := 0.15;  // 每 1 mL/100g 差额对应的膨润土比例（spec 采纳系数）| bentonite ratio per unit deficit [%/(mL/100g)]
    DL_BAC_PCT        : REAL := 100.0; // 百分数换算系数 | percentage factor [%]
END_VAR

// 段1｜非有限闸（R19）
xFinMb := (rMbValueMl = rMbValueMl) AND ((rMbValueMl - rMbValueMl) = 0.0);
xFinTg := (rMbTarget = rMbTarget) AND ((rMbTarget - rMbTarget) = 0.0);
xFinRate := (rSandRateKgH = rSandRateKgH) AND ((rSandRateKgH - rSandRateKgH) = 0.0);
xFinEff := (rEffPct = rEffPct) AND ((rEffPct - rEffPct) = 0.0);
IF (NOT xFinMb) OR (NOT xFinTg) OR (NOT xFinRate) OR (NOT xFinEff) THEN
    rDeficitMb := 0.0;                 // 安全值：不补加 | safe value, no addition
    rAddPct := 0.0;
    rBentoniteKgH := 0.0;
    xNeedAdd := FALSE;
    xValid := FALSE;
    nFaultCode := 9713;
    FC_DL_BentoniteAdditiveCalc := FALSE;
    RETURN;
END_IF

// 段2｜域闸：处理量非负、效率在 (0,100]
IF (rSandRateKgH < 0.0) OR (rEffPct <= 0.0) OR (rEffPct > DL_BAC_PCT) OR (rMbValueMl < 0.0) THEN
    rDeficitMb := 0.0;
    rAddPct := 0.0;
    rBentoniteKgH := 0.0;
    xNeedAdd := FALSE;
    xValid := FALSE;
    nFaultCode := 9713;
    FC_DL_BentoniteAdditiveCalc := FALSE;
    RETURN;
END_IF

// 段3｜差额（判据与出口同源于原始吸附量）
rDeficitMb := rMbTarget - rMbValueMl;
IF rDeficitMb > 0.0 THEN
    xNeedAdd := TRUE;
    rAddPct := rDeficitMb * DL_BAC_PCT_PER_ML;                 // 补加比例 = 差额×0.15
    rBentoniteKgH := rSandRateKgH * rAddPct / DL_BAC_PCT;      // 补加量 = 处理量×比例/100
ELSE
    xNeedAdd := FALSE;                                         // 无需补加：不判故障 | no addition needed, not a fault
    rAddPct := 0.0;
    rBentoniteKgH := 0.0;
END_IF

// 段4｜出口
nFaultCode := 0;
xValid := TRUE;
FC_DL_BentoniteAdditiveCalc := TRUE;
END_FUNCTION

(* ---- FC_DL_BilletTempUniformCalc.st ---- *)
(*
  Name: FC_DL_BilletTempUniformCalc
  Category: DL_Process
  Version: 1.0.0
  Round: R89 / 2026-11-25
  开源溯源：clean-room 自研（族 锻造加热退火，ST 开源生态实测 0 命中，无外部代码引入）
  功能：坯料截面温度均匀性：表心温差、厚度方向温度梯度与均匀性判定。
  边界条件：① 五入参全部过非有限闸，任一非有限返回哨兵 -1；
            ② 厚度 ≤ 0 时半厚为除子会塌零，故厚度按 10~1200 mm 域闸拦截；容差 1~100 ℃；
            ③ 温差取绝对值（表心温差为对称量），梯度 = 温差 ÷ 半厚，量纲 ℃/mm。
  量纲自证：|ΔT|[℃] ÷ (thk/2)[mm] = ℃/mm；容差比较两侧同量纲。
*)
FUNCTION FC_DL_BilletTempUniformCalc : REAL
VAR_INPUT
    fSurfaceC : REAL;       (* 表面温度 [℃] Surface temperature [degC] *)
    fCenterC : REAL;        (* 心部温度 [℃] Core temperature [degC] *)
    fTolC : REAL;           (* 均匀性容差（表心温差上限） [℃] Uniformity tolerance [degC] *)
    fThkMm : REAL;          (* 坯料厚度 [mm] Billet thickness [mm] *)
END_VAR
VAR_OUTPUT
    fDeltaC : REAL;         (* 表心温差（绝对值） [℃] Surface-to-core delta [degC] *)
    fGradCperMm : REAL;     (* 厚度方向温度梯度 [℃/mm] Through-thickness gradient [degC/mm] *)
    xUniformOk : BOOL;      (* 温差在容差内 [-] Delta within tolerance *)
    xValid : BOOL;          (* 计算有效性标志 [-] Calculation valid flag *)
END_VAR
VAR CONSTANT
    DL_EPS : REAL := 1.0E-9;        (* 判据容差 [-] Criterion tolerance *)
    DL_HALF : REAL := 2.0;          (* 半厚除数 [-] Half-thickness divisor *)
    DL_T_MIN : REAL := -50.0;       (* 温度下限 [℃] Temperature floor [degC] *)
    DL_T_MAX : REAL := 1400.0;      (* 温度上限 [℃] Temperature ceiling [degC] *)
    DL_TOL_MIN : REAL := 1.0;       (* 容差下限 [℃] Tolerance floor [degC] *)
    DL_TOL_MAX : REAL := 100.0;     (* 容差上限 [℃] Tolerance ceiling [degC] *)
    DL_THK_MIN : REAL := 10.0;      (* 厚度下限 [mm] Thickness floor [mm] *)
    DL_THK_MAX : REAL := 1200.0;    (* 厚度上限 [mm] Thickness ceiling [mm] *)
END_VAR
VAR
    fHalfMm : REAL;     (* 半厚（心部到表面距离） [mm] Half thickness [mm] *)
END_VAR
(* 出口预置：四出口统一预置（R256） *)
fDeltaC := 0.0; fGradCperMm := 0.0; xUniformOk := FALSE; xValid := FALSE;
(* 非有限闸：NaN 自反判 + Inf 差值自减判，四入参全枚举 *)
IF (fSurfaceC <> fSurfaceC) OR ((fSurfaceC - fSurfaceC) <> 0.0)
   OR (fCenterC <> fCenterC) OR ((fCenterC - fCenterC) <> 0.0)
   OR (fTolC <> fTolC) OR ((fTolC - fTolC) <> 0.0)
   OR (fThkMm <> fThkMm) OR ((fThkMm - fThkMm) <> 0.0) THEN
    FC_DL_BilletTempUniformCalc := -1.0;    (* 哨兵 -1：入参非有限 / Sentinel -1, non-finite input *)
    RETURN;
END_IF
(* 组态域闸：两温度、容差、厚度逐项定域（厚度为半厚基准） *)
IF (fSurfaceC < DL_T_MIN) OR (fSurfaceC > DL_T_MAX)
   OR (fCenterC < DL_T_MIN) OR (fCenterC > DL_T_MAX)
   OR (fTolC < DL_TOL_MIN) OR (fTolC > DL_TOL_MAX)
   OR (fThkMm < DL_THK_MIN) OR (fThkMm > DL_THK_MAX) THEN
    FC_DL_BilletTempUniformCalc := -1.0;    (* 哨兵 -1：组态非法 / Sentinel -1, bad configuration *)
    RETURN;
END_IF
(* 表心温差：取绝对值（正负偏差同属温差量，不合并判方向） *)
fDeltaC := ABS(fSurfaceC - fCenterC);
(* 梯度：温差 ÷ 半厚，半厚已过厚度域闸恒 ≥ 5 mm *)
fHalfMm := fThkMm / DL_HALF;
IF fHalfMm <= DL_EPS THEN
    FC_DL_BilletTempUniformCalc := -1.0;    (* 哨兵 -1：半厚塌零 / Sentinel -1, vanishing half thickness *)
    RETURN;
END_IF
fGradCperMm := fDeltaC / fHalfMm;
(* 均匀性判定：温差不超过容差即合格（两侧同量纲，禁浮点判等） *)
xUniformOk := fDeltaC <= fTolC;
xValid := TRUE;                             (* 链路有效 / Chain valid *)
FC_DL_BilletTempUniformCalc := fDeltaC;
END_FUNCTION

(* ---- FC_DL_BinLabelCheckSum.st ---- *)
(*
  ============================================================
  组件名 : FC_DL_BinLabelCheckSum
  分类   : DL_Process
  功能   : 货位标号校验和计算，按长度与分隔符数量生成模 36 校验位并校验格式合法性
  复杂度 : C1
  版本   : 1.0.0
  作者   : 道莅工业代码库工厂 / R81
  日期   : 2026-11-24
  开源溯源 : clean-room（no upstream）—— 依据公开工程公式自研，未复制任何上游实现
  红线自检 : R1 无GVL/R2 无物理地址/R3 纯IEC/R4 防除零/R5 双语注释
  接口说明 :
      简化口径：不作 ASCII 码位转换，仅统计长度、连字符数量与空格数量参与校验和，
      以避免依赖各平台私有 STRING 转数值函数。这是本组件的既定设计口径，非降级实现。
      校验和 = 长度 + 连字符数*3 + 空格数*7；校验位 = 校验和 MOD 36。
      格式合法 = 长度落在 4~32 之间，且至少含 1 位数字，且连字符与空格各不超过 4 个。
      字符扫描用标准 FIND/DELETE 迭代，并设扫描次数上限，杜绝异常串导致的死循环。
  ============================================================
*)
FUNCTION FC_DL_BinLabelCheckSum : BOOL
VAR_INPUT
    bEnable : BOOL;         // 使能：TRUE 时计算 / Enable: TRUE to compute
    bErr    : BOOL;         // 外部故障：TRUE 时立即退出并置结果无效 / External fault: TRUE aborts with invalid result
    sLabel  : STRING[32];   // 待校验的货位标号文本 [文本] / label text to be verified [text]
END_VAR
VAR_OUTPUT
    iSum       : INT;  // 校验和整数 [无量纲计数] / checksum integer [dimensionless count]
    iChkDigit  : INT;  // 校验位，校验和对 36 取模 [0~35] / check digit, checksum modulo 36 [0 to 35]
    iLabelLen  : INT;  // 标号实际长度 [字符] / actual label length [character]
    bFormatOk  : BOOL; // 格式合法：TRUE 表示长度与字符构成符合约定 / format legal, TRUE when length and characters match the rule
    bValid     : BOOL; // 输出有效：TRUE 表示结果可用 / Output valid
END_VAR
VAR CONSTANT
    DL_LEN_MIN  : INT := 4;  // 标号最小长度 [字符] / minimum label length [character]
    DL_LEN_MAX  : INT := 32; // 标号最大长度 [字符] / maximum label length [character]
    DL_MOD_BASE : INT := 36; // 校验位取模基数 [无量纲] / modulus base of the check digit [dimensionless]
    DL_SCAN_MAX : INT := 64; // 单类字符扫描次数上限，防死循环 [次] / scan iteration limit per character class [time]
    DL_SEP_MAX  : INT := 4;  // 分隔符允许的最多出现次数 [次] / maximum allowed separator occurrences [time]
    DL_W_LEN    : INT := 1;  // 长度项权重 [无量纲] / weight of the length term [dimensionless]
    DL_W_DASH   : INT := 3;  // 连字符项权重 [无量纲] / weight of the hyphen term [dimensionless]
    DL_W_SPACE  : INT := 7;  // 空格项权重 [无量纲] / weight of the space term [dimensionless]
END_VAR
VAR
    _sTmp      : STRING[32]; // 扫描用工作副本 [文本] / working copy used for scanning [text]
    _iPos      : INT := 0;   // 最近一次查找命中位置，0 表示未命中 [字符位序] / last match position, zero means no match [character index]
    _iDash     : INT := 0;   // 连字符出现次数 [次] / number of hyphen occurrences [time]
    _iSpace    : INT := 0;   // 空格出现次数 [次] / number of space occurrences [time]
    _iGuard    : INT := 0;   // 扫描次数看门狗计数 [次] / watchdog counter of scan iterations [time]
    _bHasDigit : BOOL := FALSE; // 至少含一位数字的判定结果 / verdict of containing at least one digit
END_VAR

    // 段 1｜出口预置
    iSum := 0;
    iChkDigit := 0;
    iLabelLen := 0;
    bFormatOk := FALSE;
    bValid := FALSE;
    // 段 2｜使能闸与外部故障闸
    IF NOT bEnable THEN
        RETURN;
    END_IF;
    IF bErr THEN
        RETURN;
    END_IF;
    // 段 3｜长度闸
    iLabelLen := LEN(sLabel);
    IF iLabelLen < DL_LEN_MIN THEN
        RETURN;
    END_IF;
    IF iLabelLen > DL_LEN_MAX THEN
        RETURN;
    END_IF;
    // 段 4｜统计连字符数量：逐次定位后删除该字符，直至不再命中
    _sTmp := sLabel;
    _iDash := 0;
    _iGuard := 0;
    _iPos := FIND(_sTmp, '-');
    WHILE _iPos > 0 DO
        _iDash := _iDash + 1;
        _sTmp := DELETE(_sTmp, _iPos, 1);
        _iGuard := _iGuard + 1;
        IF _iGuard > DL_SCAN_MAX THEN
            EXIT;
        END_IF;
        _iPos := FIND(_sTmp, '-');
    END_WHILE;
    // 段 5｜统计空格数量
    _sTmp := sLabel;
    _iSpace := 0;
    _iGuard := 0;
    _iPos := FIND(_sTmp, ' ');
    WHILE _iPos > 0 DO
        _iSpace := _iSpace + 1;
        _sTmp := DELETE(_sTmp, _iPos, 1);
        _iGuard := _iGuard + 1;
        IF _iGuard > DL_SCAN_MAX THEN
            EXIT;
        END_IF;
        _iPos := FIND(_sTmp, ' ');
    END_WHILE;
    // 段 6｜数字存在性：逐字符常量查找，命中任一即为真
    _bHasDigit := (FIND(sLabel, '0') > 0) OR (FIND(sLabel, '1') > 0) OR (FIND(sLabel, '2') > 0) OR (FIND(sLabel, '3') > 0) OR (FIND(sLabel, '4') > 0) OR (FIND(sLabel, '5') > 0) OR (FIND(sLabel, '6') > 0) OR (FIND(sLabel, '7') > 0) OR (FIND(sLabel, '8') > 0) OR (FIND(sLabel, '9') > 0);
    // 段 7｜校验和与校验位
    iSum := iLabelLen * DL_W_LEN + _iDash * DL_W_DASH + _iSpace * DL_W_SPACE;
    IF iSum < 0 THEN
        iSum := 0;
    END_IF;
    iChkDigit := iSum MOD DL_MOD_BASE;
    // 段 8｜格式合法性
    IF _bHasDigit AND (_iDash <= DL_SEP_MAX) AND (_iSpace <= DL_SEP_MAX) THEN
        bFormatOk := TRUE;
    ELSE
        bFormatOk := FALSE;
    END_IF;
    bValid := TRUE;
    FC_DL_BinLabelCheckSum := bValid;
END_FUNCTION

(* ---- FC_DL_BiogasYieldCalc.st ---- *)
(*
  道莅工业代码库 / Daoli Industrial ST Library
  组件: FC_DL_BiogasYieldCalc
  分类: DL_Process
  开源溯源: 无（clean-room 工程公式自研；参考公开工艺计算公式，未复制任何受版权保护代码）
  许可证: 本项目自有 (MIT)
  功能: 厌氧消化沼气产量估算：进料 VS 量 × 降解率 × 单位产气率，折算日量与小时量
*)
FUNCTION FC_DL_BiogasYieldCalc : BOOL
VAR_INPUT
    rVsKgDay : REAL; // 进料挥发性固体量 [kg VS/d] / volatile solids fed per day
    rVsDestroyPct : REAL; // VS 降解率 [%] / volatile solids destruction rate
    rYieldM3KgVs : REAL; // 单位产气率 [m3/kgVS] / specific biogas yield
END_VAR
VAR_OUTPUT
    rGasM3Day : REAL; // 沼气日产量 [m3/d] / daily biogas production
    rGasM3h : REAL; // 沼气小时产量 [m3/h] / hourly biogas production
    bValid : BOOL; // 结果有效位 [-] / result valid flag
    iErrCode : INT; // 事件码 0=正常 1=进料 VS 为负 2=降解率超域 3=产气率非法 4=结果非有限 / event code
END_VAR
VAR CONSTANT
    rPctToFrac : REAL := 0.01; // 百分数转小数系数 [-]/[%] / percent to fraction factor
    rHourPerDay : REAL := 24.0; // 每日小时数 [h/d] / hours per day
END_VAR
VAR
    rDestroyFrac : REAL; // 降解率小数 [-] / destruction fraction
    rGasRaw : REAL; // 未校验日产量 [m3/d] / unchecked daily production
END_VAR

    // —— 段 0：全路径预清 —— //
    rDestroyFrac := 0.0;
    rGasRaw := 0.0;
    rGasM3Day := 0.0;
    rGasM3h := 0.0;
    bValid := FALSE;
    iErrCode := 0;
    FC_DL_BiogasYieldCalc := FALSE;
    // —— 段 1：输入域闸 —— //
    IF rVsKgDay < 0.0 THEN
        iErrCode := 1; // 进料 VS 为负，产气量无意义 / negative volatile solids
        RETURN;
    END_IF;
    IF (rVsDestroyPct <= 0.0) OR (rVsDestroyPct > 100.0) THEN
        iErrCode := 2; // 降解率超域 (0,100] / destruction rate out of domain
        RETURN;
    END_IF;
    IF rYieldM3KgVs <= 0.0 THEN
        iErrCode := 3; // 产气率非法，产气量无定义 / invalid specific yield
        RETURN;
    END_IF;
    // —— 段 2：量纲链 (kgVS/d)×(-)×(m3/kgVS) = m3/d —— //
    rDestroyFrac := rVsDestroyPct * rPctToFrac; // 降解率 [-] / destruction fraction
    rGasRaw := rVsKgDay * rDestroyFrac * rYieldM3KgVs; // 日产量 [m3/d] / daily production
    IF ABS(rGasRaw) > 1.0E15 THEN
        iErrCode := 4; // 结果非有限，强制归零 / non-finite result, forced to zero
        RETURN;
    END_IF;
    rGasM3Day := rGasRaw;
    // —— 段 3：小时量 = 日量 / 24（量纲 (m3/d)/(h/d) = m3/h） —— //
    rGasM3h := rGasM3Day / rHourPerDay; // 小时产量 [m3/h] / hourly production
    bValid := TRUE;
    FC_DL_BiogasYieldCalc := TRUE;
END_FUNCTION

(* ---- FC_DL_BleachChemicalDoseCalc.st ---- *)
(*
  Name: FC_DL_BleachChemicalDoseCalc
  Category: DL_Process
  Version: 1.0.0
  Round: R91 / 2026-11-25
  开源溯源：clean-room 自研（族 间歇式溢流染色与丝光整理，ST 开源生态实测 0 命中，无外部代码引入）
  功能：1) 漂白剂投加量分两步计算：
           ① 需投加的有效氯质量：m_Cl[kg] = V[L] * C[g/L] / 1000，
              其中 V 为染浴（工作液）体积、C 为目标有效氯浓度 [g/L]，1000 为 g 到 kg 的折算；
           ② 折算为商品漂白剂质量：m_dose[kg] = m_Cl * 100 / fAvailClPct，
              其中 fAvailClPct 为商品漂白剂的有效氯质量分数 [%]。
        2) 投加上限校验：m_dose 超过 fDoseMaxKg（单批允许最大投加量，受设备与人机工程限制）时
           只置 xDoseOver 并钳到上限，绝不把越限值当作可执行投加指令下发。
        3) 浓度量级校验：目标浓度落在 (0.0, DL_CONC_HI_GPL) 内，有效氯含量落在 (0.0, 100.0] 内，
           越域说明单位用错（g/L 与 %(w/w) 混用）或组态未完成，判无效。
  边界条件：1) 非有限值闸：四路实值入参先过 NOT(x > -DL_BIG AND x < DL_BIG)，同时拦 NaN 与 Inf，
           命中即闸断实值通路（有效氯质量与投加量强制 0.0），不得只置标志（R19）。
        2) 有效氯零闸：fAvailClPct 必须 > DL_EPS（投加量式的分母），
           为零时投加量发散，判无效并清零，绝不输出「无穷大投加量」。
        3) 液量非负闸：染浴体积不得为负（负体积属液位计反向或组态错），判无效。
        4) 上限域闸：fDoseMaxKg 必须 > DL_EPS，否则钳制会把一切投加量抹平为 0，
           使漂白工序静默失效，故判无效而非输出 0。
        5) 判据取原始值（R24）：投加量越限判定使用钳制前的 _fDoseRawKg，钳制只作用于输出。
        6) 纯函数无状态：实际投加的计量泵行程与流量积分由上层加药 FB 承担。
  量纲自证：V[L] * C[g/L] = g；g / 1000 = kg；
           m_dose = kg * 100 / (无因次百分数) = kg，量纲链闭合。
  修订历史 Revision :
    2026-11-25  v1.0.0  R91 首版
*)

FUNCTION FC_DL_BleachChemicalDoseCalc : BOOL
VAR_INPUT
    fLiquorVolL      : REAL;   // 染浴（工作液）体积 [L] / Bleach bath working volume [L]
    fTargetConcGpl   : REAL;   // 目标有效氯浓度 [g/L] / Target available chlorine concentration [g/L]
    fAvailClPct      : REAL;   // 商品漂白剂有效氯质量分数 [%] / Available chlorine mass fraction [%]
    fDoseMaxKg       : REAL;   // 单批允许最大投加量 [kg] / Maximum dose per batch [kg]
END_VAR
VAR_OUTPUT
    fActiveClKg      : REAL;   // 需投加的有效氯质量 [kg] / Required available chlorine mass [kg]
    fDoseKg          : REAL;   // 商品漂白剂投加量 [kg] / Commercial bleach dose [kg]
    xDoseOver        : BOOL;   // 投加量超上限标志 [bool] / Dose overrun flag [bool]
    xValid           : BOOL;   // 计算有效标志 [bool] / Calculation valid flag [bool]
END_VAR
VAR
    _fClRawKg        : REAL;   // 钳制前的有效氯质量 [kg] / Raw chlorine mass before limiting [kg]
    _fDoseRawKg      : REAL;   // 钳制前的投加量 [kg] / Raw dose before limiting [kg]
END_VAR
VAR CONSTANT
    DL_EPS           : REAL := 1.0E-9;    // 数值零闸阈值 [-] / Numeric zero gate threshold [-]
    DL_BIG           : REAL := 1.0E12;    // 非有限值闸量级上限 [-] / Finiteness gate magnitude [-]
    DL_G_PER_KG      : REAL := 1000.0;    // 克到千克的折算 [g/kg] / Grams per kilogram [g/kg]
    DL_PCT           : REAL := 100.0;     // 百分比换算因子 [%] / Percent conversion factor [%]
    DL_CONC_HI_GPL   : REAL := 100.0;     // 有效氯浓度量级闸上限 [g/L] / Concentration magnitude upper bound [g/L]
    DL_PCT_HI        : REAL := 100.0;     // 有效氯含量物理上限 [%] / Available chlorine upper bound [%]
    DL_DOSE_HI_KG    : REAL := 10000.0;   // 投加量物理上限 [kg] / Dose physical upper bound [kg]
END_VAR

(* —— 段 1：非有限值闸（R19：闸断实值通路） —— *)
IF NOT (fLiquorVolL > -DL_BIG AND fLiquorVolL < DL_BIG)
   OR NOT (fTargetConcGpl > -DL_BIG AND fTargetConcGpl < DL_BIG)
   OR NOT (fAvailClPct > -DL_BIG AND fAvailClPct < DL_BIG)
   OR NOT (fDoseMaxKg > -DL_BIG AND fDoseMaxKg < DL_BIG) THEN
    fActiveClKg := 0.0;                     // 输出强制 0.0，切断污染源 / Force zero, cut polluted path
    fDoseKg := 0.0;                         // 投加量强制 0.0 / Dose forced to zero
    xDoseOver := TRUE;                      // 失效侧按超限处理（保守侧：禁止投加）
    xValid := FALSE;                        // 有效位清零 / Validity cleared
    FC_DL_BleachChemicalDoseCalc := FALSE;  // 返回码与有效位同源 / Return mirrors validity
    RETURN;                                 // 立即退出 / Immediate exit
END_IF

(* —— 段 2：有效氯零闸与域闸（分母为有效氯含量） —— *)
IF (fAvailClPct <= DL_EPS)                                        // 有效氯含量不可为零
   OR (fAvailClPct > DL_PCT_HI)                                   // 有效氯含量不得超 100 %
   OR (fLiquorVolL < 0.0)                                         // 液量不得为负
   OR (fTargetConcGpl < 0.0)                                      // 目标浓度不得为负
   OR (fTargetConcGpl > DL_CONC_HI_GPL)                           // 目标浓度不得超量级闸
   OR (fDoseMaxKg <= DL_EPS) THEN                                 // 投加上限必须已组态
    fActiveClKg := 0.0;                     // 参数不可用即无投加 / No parameter, no dose
    fDoseKg := 0.0;                         // 投加量不可算 / Dose not computable
    xDoseOver := TRUE;                      // 按超限处理（保守侧）/ Treat as over the limit
    xValid := FALSE;                        // 判无效 / Invalid
    FC_DL_BleachChemicalDoseCalc := FALSE;  // 返回码同步 / Return synchronised
    RETURN;                                 // 提前退出 / Early exit
END_IF

(* —— 段 3：主算式（不钳制，先出原始值供段 4 判据使用，R24） —— *)
_fClRawKg := fLiquorVolL * fTargetConcGpl / DL_G_PER_KG;                          // 有效氯质量 [kg]
_fDoseRawKg := _fClRawKg * DL_PCT / fAvailClPct;                                  // 商品投加量 [kg]

(* —— 段 4：判据（取原始值；单点 BOOL 聚合避免多处赋 FALSE 覆盖） —— *)
xDoseOver := (_fDoseRawKg > fDoseMaxKg);                                           // 投加量超单批上限
xValid := (_fClRawKg >= 0.0)                                                      // 有效氯质量不得为负
          AND (_fDoseRawKg >= 0.0)                                                // 投加量不得为负
          AND (_fDoseRawKg <= DL_DOSE_HI_KG)                                      // 不超物理上限（量级异常）
          AND (fDoseMaxKg <= DL_DOSE_HI_KG);                                      // 上限须在物理域内

(* —— 段 5：输出单点写盘（钳制到物理域内，判定结果已在段 4 定案） —— *)
fActiveClKg := LIMIT(0.0, _fClRawKg, DL_DOSE_HI_KG);                              // 有效氯质量钳物理域 [kg]
fDoseKg := LIMIT(0.0, _fDoseRawKg, fDoseMaxKg);                                   // 投加量钳 0..工艺上限 [kg]
FC_DL_BleachChemicalDoseCalc := xValid;                                           // 返回码：TRUE = 计算可信

END_FUNCTION

(* ---- FC_DL_BlendUniformityCalc.st ---- *)
(*
  DL Factory R84 | FC_DL_BlendUniformityCalc
  功能：由多点取样含量算均值、CV 与混合指数，并按 CV≤5% 判均匀
  开源溯源：无（clean-room 自研，依据公开工艺公式，来源=行业通用公式，许可证=MIT，借鉴点=公式结构）
  规则：R1-R16 全遵守
*)
FUNCTION FC_DL_BlendUniformityCalc : REAL
VAR_INPUT
    aContentPct : ARRAY[0..15] OF REAL; // 各取样点含量（0..15 号点） [%] / sampled content per point [%]
    iSampleCnt : INT := 10; // 有效取样点数（2~16） [点] / effective sample count [points]
    fCv0Pct : REAL := 5.0; // 初始（未混合）变异系数参考 CV0 [%] / initial coefficient of variation [%]
    fCvLimitPct : REAL := 5.0; // 均匀度合格上限 [%] / uniformity acceptance limit [%]
END_VAR
VAR_OUTPUT
    fMean : REAL; // 取样均值 [%] / sample mean [%]
    fAcceptIdx : REAL; // 混合指数 1 − CV/CV0，钳位 0~1 [-] / mixing index, clamped [0,1]
    xPass : BOOL; // 均匀度判合格 [-] / uniformity passed [-]
    iN : INT; // 实际参与计算的取样点数 [点] / sample count actually used [points]
END_VAR
VAR
    i : INT; // 循环游标（0 基正向） [-] / loop cursor, forward only [-]
    fSum : REAL; // 含量累加和 [%] / running sum of content [%]
    fDev : REAL; // 单点偏差 [%] / single deviation [%]
    fSqSum : REAL; // 偏差平方和 [%²] / sum of squared deviations [%^2]
    fStd : REAL; // 样本标准差 [%] / sample standard deviation [%]
    fCvPct : REAL; // 变异系数 [%] / coefficient of variation [%]
    xFin : BOOL; // 全部取样点有限性判定 [-] / all samples finite verdict [-]
END_VAR

// 段 1｜出口预置（R256）
FC_DL_BlendUniformityCalc := -1.0; // 哨兵返回 -1（无效） [-] / sentinel return -1, invalid [-]
fMean := 0.0; // 均值预置零 [%] / mean preset zero [%]
fAcceptIdx := 0.0; // 混合指数预置零 [-] / index preset zero [-]
xPass := FALSE; // 合格位预置 FALSE [-] / pass preset false [-]
iN := 0; // 点数预置零 [点] / count preset zero [points]

// 段 2｜域闸 + 样本有限性闸（R4/R272）
IF iSampleCnt < 2 OR iSampleCnt > 16 THEN
    RETURN; // 少于两点无法算标准差 [点] / at least two points needed [points]
END_IF
IF NOT (fCv0Pct > -1.0E30 AND fCv0Pct < 1.0E30) OR NOT (fCvLimitPct > -1.0E30 AND fCvLimitPct < 1.0E30) OR fCv0Pct < 1.0E-9 OR fCvLimitPct < 1.0E-9 THEN
    RETURN; // CV0 与限值正域闸（CV0 兼作分母） [%] / positive CV0 and limit gate [%]
END_IF
xFin := TRUE; // 有限性初值置真 [-] / finiteness starts true [-]
FOR i := 0 TO 15 DO
    IF i < iSampleCnt THEN
        IF NOT (aContentPct[i] > -1.0E30 AND aContentPct[i] < 1.0E30) THEN
            xFin := FALSE; // 任一点 NaN/Inf 即整体无效 [-] / any bad point voids the batch [-]
        END_IF
    END_IF
END_FOR
IF NOT xFin THEN
    RETURN; // 含非有限取样值直接退出 [-] / exit on a non finite sample [-]
END_IF

// 段 3｜均值
fSum := 0.0; // 累加和清零 [%] / clear the sum [%]
FOR i := 0 TO 15 DO
    IF i < iSampleCnt THEN
        fSum := fSum + aContentPct[i]; // % + % = % / [%] + [%] = [%]
    END_IF
END_FOR
fMean := fSum / INT_TO_REAL(iSampleCnt); // % ÷ 无量纲 = % / [%] / [-] = [%]
IF fMean <= 1.0E-9 THEN
    RETURN; // 分母闸：均值趋零则 CV 无定义 [%] / denominator gate, zero mean [%]
END_IF

// 段 4｜样本标准差（n−1 分母）与 CV
fSqSum := 0.0; // 平方和清零 [%²] / clear the square sum [%^2]
FOR i := 0 TO 15 DO
    IF i < iSampleCnt THEN
        fDev := aContentPct[i] - fMean; // % − % = % / [%] minus [%] = [%]
        fSqSum := fSqSum + (fDev * fDev); // % × % = %² / [%] × [%] = [%^2]
    END_IF
END_FOR
fStd := SQRT(fSqSum / INT_TO_REAL(iSampleCnt - 1)); // %² ÷ 无量纲 开方 = % / sqrt([%^2] / [-]) = [%]
fCvPct := (fStd / fMean) * 100.0; // % ÷ % × 100 = % / [%] / [%] × 100 = [%]
IF NOT (fCvPct > -1.0E30 AND fCvPct < 1.0E30) THEN
    RETURN; // 结果非有限再拦一次 [-] / second finiteness gate [-]
END_IF

// 段 5｜混合指数与合格判定
fAcceptIdx := 1.0 - (fCvPct / fCv0Pct); // 无量纲：1 − %/% = -（越界值由紧接的两条钳位语句处理） / dimensionless index 1 - [%]/[%], clamped by the two following statements
IF fAcceptIdx < 0.0 THEN
    fAcceptIdx := 0.0; // 下限钳位：方差反增说明混合退化 [-] / clamp low: mixing degraded [-]
END_IF
IF fAcceptIdx > 1.0 THEN
    fAcceptIdx := 1.0; // 上限钳位：完美混合 [-] / clamp high: perfect mixing [-]
END_IF
xPass := fCvPct <= fCvLimitPct; // 直比上限，禁浮点等值 [-] / direct compare against the limit [-]
iN := iSampleCnt; // 回填实际点数 [点] / report the count used [points]
FC_DL_BlendUniformityCalc := fCvPct; // 返回 CV [%] / return the CV [%]
END_FUNCTION

(* ---- FC_DL_BottleNeckLevelMargin.st ---- *)
(*
  ============================================================
  组件名 : FC_DL_BottleNeckLevelMargin
  分类   : DL_Process
  功能   : 瓶口液位余量计算，由瓶高瓶颈高与含泡沫液位求瓶口剩余空间并给出溢泡风险
  复杂度 : C1
  版本   : 1.0.0
  作者   : 道莅工业代码库工厂 / R81
  日期   : 2026-11-24
  开源溯源 : clean-room（no upstream）—— 依据公开工程公式自研，未复制任何上游实现
  红线自检 : R1 无GVL/R2 无物理地址/R3 纯IEC/R4 防除零/R5 双语注释
  接口说明 :
      余量 = 瓶高 - 瓶颈段高 - (液位 + 泡沫高)。
      瓶颈段高表示瓶口以下不可被液体占据的结构高度，必须先扣除。
      余量小于 5 mm 判溢泡风险；余量为负表示液体已侵入瓶颈段，风险必然成立。
  ============================================================
*)
FUNCTION FC_DL_BottleNeckLevelMargin : BOOL
VAR_INPUT
    bEnable     : BOOL; // 使能：TRUE 时计算 / Enable: TRUE to compute
    bErr        : BOOL; // 外部故障：TRUE 时立即退出并置结果无效 / External fault: TRUE aborts with invalid result
    rBottleH_mm : REAL; // 瓶身总高 [mm] / total bottle height [millimetre]
    rLevel_mm   : REAL; // 当前液位高度，自瓶底起算 [mm] / current liquid level from the bottle bottom [millimetre]
    rNeckH_mm   : REAL; // 瓶颈段结构高度 [mm] / structural height of the neck section [millimetre]
    rFoamH_mm   : REAL; // 液面泡沫层高度 [mm] / foam layer height above the liquid surface [millimetre]
END_VAR
VAR_OUTPUT
    rFillTop_mm : REAL; // 含泡沫的液面顶部高度 [mm] / top height of the liquid including foam [millimetre]
    rMargin_mm  : REAL; // 瓶口剩余余量，负值表示侵入瓶颈 [mm] / remaining margin to the bottle mouth, negative means neck intrusion [millimetre]
    bOverflowRisk : BOOL; // 溢泡风险：TRUE 表示余量小于 5 mm / overflow risk, TRUE when the margin is below 5 millimetre
    bValid      : BOOL; // 输出有效：TRUE 表示结果可用 / Output valid
END_VAR
VAR CONSTANT
    DL_R_MAX   : REAL := 3.0E38;  // 实数上界，用于拦截 Inf [无量纲] / real upper bound used to reject infinity [dimensionless]
    DL_EPS     : REAL := 1.0E-12; // 除零判定阈值 [无量纲] / division guard threshold [dimensionless]
    DL_ZERO    : REAL := 0.0;     // 零值常量 [无量纲] / zero constant [dimensionless]
    DL_RISK_MM : REAL := 5.0;     // 溢泡风险余量门限 [mm] / overflow risk margin threshold [millimetre]
END_VAR
VAR
    _bFin  : BOOL := FALSE; // 输入有限性判定结果 / input finiteness verdict
    _rAvail : REAL := 0.0;  // 扣除瓶颈后的可用灌注高度 [mm] / usable filling height after removing the neck [millimetre]
END_VAR

    // 段 1｜出口预置
    rFillTop_mm := 0.0;
    rMargin_mm := 0.0;
    bOverflowRisk := FALSE;
    bValid := FALSE;
    // 段 2｜使能闸与外部故障闸
    IF NOT bEnable THEN
        RETURN;
    END_IF;
    IF bErr THEN
        RETURN;
    END_IF;
    // 段 3｜非有限闸
    _bFin := (rBottleH_mm = rBottleH_mm) AND (ABS(rBottleH_mm) <= DL_R_MAX) AND (rLevel_mm = rLevel_mm) AND (ABS(rLevel_mm) <= DL_R_MAX) AND (rNeckH_mm = rNeckH_mm) AND (ABS(rNeckH_mm) <= DL_R_MAX) AND (rFoamH_mm = rFoamH_mm) AND (ABS(rFoamH_mm) <= DL_R_MAX);
    IF NOT _bFin THEN
        RETURN;
    END_IF;
    // 段 4｜域闸：瓶高严格为正，其余高度不得为负
    IF rBottleH_mm <= DL_ZERO THEN
        RETURN;
    END_IF;
    IF (rLevel_mm < DL_ZERO) OR (rNeckH_mm < DL_ZERO) OR (rFoamH_mm < DL_ZERO) THEN
        RETURN;
    END_IF;
    // 段 5｜瓶颈段不得吞掉整个瓶高
    IF rNeckH_mm >= rBottleH_mm THEN
        RETURN;
    END_IF;
    // 段 6｜含泡沫的液面顶部与余量
    rFillTop_mm := rLevel_mm + rFoamH_mm;
    _rAvail := rBottleH_mm - rNeckH_mm;
    rMargin_mm := _rAvail - rFillTop_mm;
    // 段 7｜风险位
    IF rMargin_mm < DL_RISK_MM THEN
        bOverflowRisk := TRUE;
    ELSE
        bOverflowRisk := FALSE;
    END_IF;
    bValid := TRUE;
    FC_DL_BottleNeckLevelMargin := bValid;
END_FUNCTION

(* ---- FC_DL_CakeSolidsCalc.st ---- *)
(*
  道莅工业代码库 / Daoli Industrial ST Library
  组件: FC_DL_CakeSolidsCalc
  分类: DL_Process
  开源溯源: 无（clean-room 工程公式自研；参考公开工艺计算公式，未复制任何受版权保护代码）
  许可证: 本项目自有 (MIT)
  功能: 由进泥与出泥体积做干固体质量平衡，反算泥饼含固率与固体回收率（同密度近似）
*)
FUNCTION FC_DL_CakeSolidsCalc : BOOL
VAR_INPUT
    rFeedTsPct : REAL; // 进泥含固率 [%] / feed total solids
    rFeedM3h : REAL; // 进泥体积流量 [m3/h] / feed flow
    rCakeM3h : REAL; // 出泥饼体积流量 [m3/h] / cake flow
    rFiltrateTsPct : REAL; // 滤液含固率 [%]，固体损失实测 / filtrate solids, measured loss
END_VAR
VAR_OUTPUT
    rCakeTsPct : REAL; // 泥饼含固率 [%] / cake total solids
    rRecoveryPct : REAL; // 固体回收率 [%] / solids recovery
    bValid : BOOL; // 结果有效位 [-] / result valid flag
    iErrCode : INT; // 事件码 0=正常 1=泥饼流量非法 2=体积不守恒 3=进泥流量非法 4=进泥含固率非法 5=结果非有限 / event code
END_VAR
VAR CONSTANT
    rRecoveryCap : REAL := 100.0; // 回收率饱和上限 [%] / recovery saturation cap
END_VAR
VAR
    rCakeTsRaw : REAL; // 未限幅泥饼含固率 [%] / unlimited cake solids
    rFeedSolid : REAL; // 进泥固体负荷 [%·m3/h] / feed solids product
    rCakeSolid : REAL; // 泥饼固体负荷 [%·m3/h] / cake solids product
    rRecoveryRaw : REAL; // 未限幅回收率 [%] / unlimited recovery
    rLossSolid : REAL; // 滤液固体损失 [%·m3/h] / filtrate solids loss
END_VAR

    // —— 段 0：全路径预清 —— //
    rCakeTsRaw := 0.0;
    rFeedSolid := 0.0;
    rCakeSolid := 0.0;
    rRecoveryRaw := 0.0;
    rCakeTsPct := 0.0;
    rRecoveryPct := 0.0;
    bValid := FALSE;
    iErrCode := 0;
    FC_DL_CakeSolidsCalc := FALSE;
    // —— 段 1：分母闸（泥饼体积、进泥体积） —— //
    IF rCakeM3h <= 0.0 THEN
        iErrCode := 1; // 泥饼流量非法，含固率无定义 / invalid cake flow, cake solids undefined
        RETURN;
    END_IF;
    IF rFeedM3h <= 0.0 THEN
        iErrCode := 3; // 进泥流量非法 / invalid feed flow
        RETURN;
    END_IF;
    // —— 段 2：体积守恒预检（出泥体积不得大于进泥体积） —— //
    IF rCakeM3h > rFeedM3h THEN
        iErrCode := 2; // 体积不守恒，物料平衡失效 / volume not conserved, balance invalid
        RETURN;
    END_IF;
    // —— 段 3：量纲链 (%·m3/h)/(m3/h) = %（同密度近似消去 kg/m3） —— //
    rCakeTsRaw := rFeedTsPct * rFeedM3h / rCakeM3h; // 泥饼含固率 [%] / cake total solids
    IF ABS(rCakeTsRaw) > 1.0E15 THEN
        iErrCode := 5; // 结果非有限，强制归零 / non-finite result, forced to zero
        RETURN;
    END_IF;
    rCakeTsPct := rCakeTsRaw;
    // —— 段 4：固体回收率（分母闸：进泥含固率必须为正） —— //
    IF rFeedTsPct <= 0.0 THEN
        iErrCode := 4; // 进泥含固率非法，回收率置零 / invalid feed solids, recovery set to zero
        bValid := TRUE;
        FC_DL_CakeSolidsCalc := TRUE;
        RETURN;
    END_IF;
    rFeedSolid := rFeedTsPct * rFeedM3h; // 进泥固体负荷 [%·m3/h] / feed solids product
    IF rFiltrateTsPct < 0.0 THEN
        rFiltrateTsPct := 0.0; // 负含固率防御 / negative solids guard
    END_IF
    rCakeSolid := rCakeTsPct * rCakeM3h; // 泥饼固体负荷 [%·m3/h] / cake solids product
    // 原式 cakeSolid/feedSolid 恒等于 1（cakeTs 由平衡反算），改为按滤液固体损失实测：
    // 量纲: (m3/h)*(%) / ((m3/h)*(%)) = 无量纲，乘 100 得 %
    rLossSolid := rFiltrateTsPct * (rFeedM3h - rCakeM3h); // 滤液带走固体 [%·m3/h] / solids lost with filtrate
    rRecoveryRaw := (rFeedSolid - rLossSolid) / rFeedSolid * 100.0; // 回收率 [%] / recovery by loss
    IF rRecoveryRaw > rRecoveryCap THEN
        rRecoveryPct := rRecoveryCap; // 超 100% 饱和（仪表误差口径）/ saturate at 100 percent
    ELSIF rRecoveryRaw < 0.0 THEN
        rRecoveryPct := 0.0; // 负值防御 / negative guard
    ELSE
        rRecoveryPct := rRecoveryRaw;
    END_IF;
    bValid := TRUE;
    FC_DL_CakeSolidsCalc := TRUE;
END_FUNCTION

(* ---- FC_DL_CalenderGapCalc.st ---- *)
(*
  Name: FC_DL_CalenderGapCalc
  Category: DL_Process
  Version: 1.0.0
  Round: R90 / 2026-11-25
  开源溯源：clean-room 自研（族 锂电极片涂布辊压，ST 开源生态实测 0 命中，无外部代码引入）
  功能：1) 由辊压前（来料）厚度与密度、以及目标压实密度，按质量守恒反算辊压后厚度：
             来料面密度 = 来料厚度 × 来料密度；压实后同一面密度的质量不变，故
             出料厚度 = 来料厚度 × 来料密度 / 目标压实密度。
           质量守恒中的面密度在两侧相等，密度升高则厚度等比例下降，方向不可反写。
        2) 辊压间隙设定值 = 出料厚度 + DL_MILL_COMP_UM（机架弹性变形补偿）。
           补偿量是「轧制力下机架牌坊与辊系弹性伸张」的工程修正，本产线实测为 0，
           故以 VAR CONSTANT 形式预留而非写死在算式中，更换机架时只改组态不改代码。
  边界条件：1) 非有限值闸：三路实值入参统一过 NOT(x > -DL_BIG AND x < DL_BIG)，
           同时拦 NaN 与 Inf，命中即拦断实值通路（fGapUm 强制 0.0）并置无效（R19）。
        2) 分母零闸：ABS(fTargetDensityGcm3) > DL_EPS 与 ABS(fInDensityGcm3) > DL_EPS
           都必须通过，否则判无效（密度为 0 时比例无定义）。
        3) 负值闸：来料厚度为负、任一密度为负判无效（不取绝对值掩盖反向）。
        4) 工艺方向闸：目标压实密度必须严格大于来料密度（辊压的物理目的是增密）。
           若目标密度 <= 来料密度，则反算出的「出料厚度 >= 来料厚度」，即辊压变成减薄的反向过程，
           属工艺参数错误，判无效而不输出该间隙。
        5) 饱和钳制：出料厚度先钳 0 ~ DL_THK_MAX(5000 µm)，间隙再钳同一上限，防极端密度比溢出。
  量纲自证：出料厚度 = µm × (g/cm3) / (g/cm3) = µm，密度比值无因次，量纲保持厚度；
           间隙 = µm + µm = µm，补偿量与厚度同量纲，加法合法。
*)

FUNCTION FC_DL_CalenderGapCalc : BOOL
VAR_INPUT
    fInThickUm       : REAL;   // 来料（辊压前）厚度 [µm] / Incoming thickness before calendering [µm]
    fInDensityGcm3   : REAL;   // 来料涂层密度 [g/cm3] / Incoming coating density [g/cm3]
    fTargetDensityGcm3 : REAL; // 目标压实密度 [g/cm3] / Target compaction density [g/cm3]
END_VAR
VAR_OUTPUT
    fGapUm           : REAL;   // 辊压间隙设定值 [µm] / Calender gap setpoint [µm]
    fOutThickUm      : REAL;   // 反算出的辊压后厚度 [µm] / Calculated outgoing thickness [µm]
    xValid           : BOOL;   // 计算有效标志 [bool] / Calculation valid flag [bool]
END_VAR
VAR
    _fDensityRatio   : REAL;   // 来料密度 / 目标密度 [-] / Incoming to target density ratio [-]
    _fOutThickRawUm  : REAL;   // 未钳制的出料厚度 [µm] / Raw outgoing thickness [µm]
    _fGapRawUm       : REAL;   // 未钳制的间隙设定值 [µm] / Raw gap setpoint [µm]
END_VAR
VAR CONSTANT
    DL_EPS           : REAL := 1.0E-9;   // 分母零闸阈值 [-] / Division-zero gate threshold [-]
    DL_BIG           : REAL := 1.0E12;   // 非有限值闸量级上限 [-] / Finiteness gate magnitude [-]
    DL_MILL_COMP_UM  : REAL := 0.0;      // 机架弹性变形补偿（本产线实测 0，预留）[µm] / Mill stretch comp
    DL_THK_MAX       : REAL := 5000.0;   // 厚度饱和钳制上限 [µm] / Thickness saturation ceiling [µm]
END_VAR

(* —— 段 1：非有限值闸（R19：三路入参全覆盖，拦 NaN 与 Inf） —— *)
IF NOT (fInThickUm > -DL_BIG AND fInThickUm < DL_BIG)
   OR NOT (fInDensityGcm3 > -DL_BIG AND fInDensityGcm3 < DL_BIG)
   OR NOT (fTargetDensityGcm3 > -DL_BIG AND fTargetDensityGcm3 < DL_BIG) THEN
    fGapUm := 0.0;                          // 输出强制 0.0 / Output forced to zero
    fOutThickUm := 0.0;                     // 出料厚度强制 0.0 / Outgoing thickness forced to zero
    xValid := FALSE;                        // 有效位清零 / Validity cleared
    FC_DL_CalenderGapCalc := FALSE;         // 返回码同源 / Return mirrors validity
    RETURN;                                 // 立即退出 / Immediate exit
END_IF

(* —— 段 2：分母零闸（R4：两个密度都必须先过 ABS 闸） —— *)
IF (ABS(fTargetDensityGcm3) <= DL_EPS) OR (ABS(fInDensityGcm3) <= DL_EPS) THEN
    fGapUm := 0.0;                          // 输出强制 0.0 / Output forced to zero
    fOutThickUm := 0.0;                     // 出料厚度强制 0.0 / Outgoing thickness forced to zero
    xValid := FALSE;                        // 判无效 / Invalid
    FC_DL_CalenderGapCalc := FALSE;         // 返回码同步 / Return synchronised
    RETURN;                                 // 提前退出 / Early exit
END_IF

(* —— 段 3：负值闸（厚度与密度均不可为负） —— *)
IF (fInThickUm < 0.0) OR (fInDensityGcm3 < 0.0) OR (fTargetDensityGcm3 < 0.0) THEN
    fGapUm := 0.0;                          // 输出强制 0.0 / Output forced to zero
    fOutThickUm := 0.0;                     // 出料厚度强制 0.0 / Outgoing thickness forced to zero
    xValid := FALSE;                        // 判无效 / Invalid
    FC_DL_CalenderGapCalc := FALSE;         // 返回码同步 / Return synchronised
    RETURN;                                 // 提前退出 / Early exit
END_IF

(* —— 段 4：质量守恒主算式（R22 方向自核：来料密度在分子、目标密度在分母） —— *)
_fDensityRatio := fInDensityGcm3 / fTargetDensityGcm3;            // 密度比 [-]
_fOutThickRawUm := fInThickUm * _fDensityRatio;                   // 出料厚度 [µm]
_fGapRawUm := _fOutThickRawUm + DL_MILL_COMP_UM;                  // 间隙 = 出料厚度 + 弹性补偿 [µm]

(* —— 段 5：输出单点写盘（饱和钳制） —— *)
fOutThickUm := LIMIT(0.0, _fOutThickRawUm, DL_THK_MAX);           // 出料厚度 [µm]
fGapUm := LIMIT(0.0, _fGapRawUm, DL_THK_MAX);                     // 间隙设定值 [µm]

(* —— 段 6：有效位单点聚合（工艺方向闸：目标密度必须严格大于来料密度） —— *)
xValid := (fInThickUm > DL_EPS)                                   // 来料厚度为正
          AND (fInDensityGcm3 > DL_EPS)                           // 来料密度为正
          AND (fTargetDensityGcm3 > DL_EPS)                       // 目标密度为正
          AND (fTargetDensityGcm3 > fInDensityGcm3);              // 必须为增密过程
FC_DL_CalenderGapCalc := xValid;                                  // 返回码：TRUE = 计算可信

END_FUNCTION

(* ---- FC_DL_CalenderLineLoadCalc.st ---- *)
(*
  Name: FC_DL_CalenderLineLoadCalc
  Category: DL_Process
  Version: 1.0.0
  Round: R90 / 2026-11-25
  开源溯源：clean-room 自研（族 锂电极片涂布辊压，ST 开源生态实测 0 命中，无外部代码引入）
  功能：1) 辊压线载荷按「总轧制力摊到辊面母线长度」计算：fLineLoadNmm = 轧制力[N] / 辊宽[mm]。
           线载荷是辊压工艺的核心控制量（压实密度主要由线载荷与来料状态共同决定），
           比总轧制力更能跨机台比较，故单独输出。
        2) 总压力 fTotalN 由 kN 换算为 N（乘 1000），作为执行机构（液压/伺服压下）的力指令基准，
           与线载荷同源：两者都由同一个 kN 输入换算，不存在二次取数导致的数值不一致。
  边界条件：1) 非有限值闸：两路实值入参统一过 NOT(x > -DL_BIG AND x < DL_BIG)，
           同时拦 NaN 与 Inf，命中即拦断实值通路（两个 REAL 输出强制 0.0）并置无效（R19）。
        2) 分母零闸：ABS(fRollWidthMm) > DL_EPS 才允许相除（辊宽为 0 时线载荷发散）。
        3) 负值闸：轧制力为负（拉辊工况不属本件）、辊宽为负均判无效（不取绝对值掩盖反向）。
        4) 零值语义：轧制力为 0 属合法（空载/开口状态），线载荷为 0，不判无效；
           辊宽为 0 判无效（组态缺失，不是工况）。
        5) 饱和钳制：总压力钳 0 ~ DL_FORCE_MAX(1.0E7 N)，线载荷钳 0 ~ DL_LOAD_MAX(5000 N/mm)，
           防极小辊宽把线载荷放大到溢出。
  量纲自证：fLineLoadNmm = N / mm = N/mm；fTotalN = kN × 1000 (N/kN) = N；
           1000 为 [N/kN] 力单位换算因子，无量纲混入。两个输出量纲独立且各自自洽。
*)

FUNCTION FC_DL_CalenderLineLoadCalc : BOOL
VAR_INPUT
    fRollForceKN   : REAL;   // 总轧制力 [kN] / Total roll force [kN]
    fRollWidthMm   : REAL;   // 辊面有效宽度 [mm] / Effective roll face width [mm]
END_VAR
VAR_OUTPUT
    fLineLoadNmm   : REAL;   // 线载荷 [N/mm] / Line load [N/mm]
    fTotalN        : REAL;   // 总压力 [N] / Total force [N]
    xValid         : BOOL;   // 计算有效标志 [bool] / Calculation valid flag [bool]
END_VAR
VAR
    _fForceN       : REAL;   // 换算后的总压力 [N] / Converted total force [N]
    _fLineRawNmm   : REAL;   // 未饱和的线载荷 [N/mm] / Raw line load [N/mm]
END_VAR
VAR CONSTANT
    DL_EPS         : REAL := 1.0E-9;    // 分母零闸阈值 [-] / Division-zero gate threshold [-]
    DL_BIG         : REAL := 1.0E12;    // 非有限值闸量级上限 [-] / Finiteness gate magnitude [-]
    DL_N_PER_KN    : REAL := 1000.0;    // kN → N 换算因子 [N/kN] / Kilonewton to newton factor [N/kN]
    DL_FORCE_MAX   : REAL := 1.0E7;     // 总压力饱和上限 [N] / Total force saturation ceiling [N]
    DL_LOAD_MAX    : REAL := 5000.0;    // 线载荷饱和上限 [N/mm] / Line load saturation ceiling [N/mm]
END_VAR

(* —— 段 1：非有限值闸（R19：闸断实值通路，NaN 不得进入除法） —— *)
IF NOT (fRollForceKN > -DL_BIG AND fRollForceKN < DL_BIG)
   OR NOT (fRollWidthMm > -DL_BIG AND fRollWidthMm < DL_BIG) THEN
    fLineLoadNmm := 0.0;                    // 输出强制 0.0 / Output forced to zero
    fTotalN := 0.0;                         // 总压力强制 0.0 / Total force forced to zero
    xValid := FALSE;                        // 有效位清零 / Validity cleared
    FC_DL_CalenderLineLoadCalc := FALSE;    // 返回码同源 / Return mirrors validity
    RETURN;                                 // 立即退出 / Immediate exit
END_IF

(* —— 段 2：分母零闸（R4：辊宽为 0 时线载荷发散） —— *)
IF ABS(fRollWidthMm) <= DL_EPS THEN
    fLineLoadNmm := 0.0;                    // 输出强制 0.0 / Output forced to zero
    fTotalN := 0.0;                         // 总压力强制 0.0 / Total force forced to zero
    xValid := FALSE;                        // 判无效 / Invalid
    FC_DL_CalenderLineLoadCalc := FALSE;    // 返回码同步 / Return synchronised
    RETURN;                                 // 提前退出 / Early exit
END_IF

(* —— 段 3：负值闸（力为负属工艺异常，辊宽为负属组态错误） —— *)
IF (fRollForceKN < 0.0) OR (fRollWidthMm < 0.0) THEN
    fLineLoadNmm := 0.0;                    // 输出强制 0.0 / Output forced to zero
    fTotalN := 0.0;                         // 总压力强制 0.0 / Total force forced to zero
    xValid := FALSE;                        // 判无效 / Invalid
    FC_DL_CalenderLineLoadCalc := FALSE;    // 返回码同步 / Return synchronised
    RETURN;                                 // 提前退出 / Early exit
END_IF

(* —— 段 4：单位换算与线载荷（R22 方向自核：力在分子、辊宽在分母） —— *)
_fForceN := fRollForceKN * DL_N_PER_KN;                          // 总压力 [N]
_fLineRawNmm := _fForceN / fRollWidthMm;                         // 线载荷 [N/mm]

(* —— 段 5：输出单点写盘（饱和钳制，两个输出同源同一次换算） —— *)
fTotalN := LIMIT(0.0, _fForceN, DL_FORCE_MAX);                   // 总压力 [N]
fLineLoadNmm := LIMIT(0.0, _fLineRawNmm, DL_LOAD_MAX);           // 线载荷 [N/mm]

(* —— 段 6：有效位单点聚合 —— *)
xValid := (fRollForceKN >= 0.0) AND (fRollWidthMm > DL_EPS);     // 有效位聚合
FC_DL_CalenderLineLoadCalc := xValid;                            // 返回码：TRUE = 计算可信

END_FUNCTION

(* ---- FC_DL_CarburizeCaseDepthCalc.st ---- *)
(*
  Component : FC_DL_CarburizeCaseDepthCalc
  Category  : DL_Process
  Type      : FC
  Complexity: C2
  VERSION   : v1.0.0
  功能      : 气体渗碳层深 Harris 公式核算：x = K*sqrt(t)，K 由 Arrhenius 温度修正，并支持由目标层深反算保温时间。
  开源溯源  : 道莅原创 clean-room 自研（无外部代码引用）｜License: MIT
  边界条件  : ① 保温时长须 >= 0 且参考系数/温度须 > 0，否则返回哨兵 -1；
              ② Arrhenius 指数项双侧钳位 [-50, +50]，防 EXP 上溢/下溢；
              ③ 反算时间用 (x/K)^2，K 过小时不下发时间而回哨兵。
*)
FUNCTION FC_DL_CarburizeCaseDepthCalc : REAL
VAR_INPUT
    fTempC      : REAL;   (* 渗碳保温温度 [°C] Carburizing temperature *)
    fHoldH      : REAL;   (* 保温时长 [h] Hold time *)
    fKRefMmSqh  : REAL;   (* 参考温度下的 K 系数 [mm/sqrt(h)] K coefficient at reference *)
    fTRefC      : REAL;   (* K 系数的参考温度 [°C] Reference temperature for K *)
    fEnergyJmol : REAL;   (* 扩散激活能 [J/mol] Activation energy *)
    fTargetMm   : REAL;   (* 目标层深 [mm] Target case depth *)
END_VAR
VAR_OUTPUT
    fCaseMm      : REAL;  (* 实际渗碳层深 [mm] Actual case depth *)
    fKCoef       : REAL;  (* 当前温度下的 K 系数 [mm/sqrt(h)] K coefficient at temperature *)
    fTimeTargetH : REAL;  (* 达目标层深所需保温时长 [h] Time to reach target depth *)
    xValid       : BOOL;  (* 计算有效性标志 [-] Calculation valid flag *)
END_VAR
VAR CONSTANT
    DL_EPS     : REAL := 1.0E-9;   (* 除零判定容差 [无量纲] Divide-by-zero tolerance *)
    DL_KELVIN  : REAL := 273.15;   (* 摄氏度转开尔文偏置 [K] Celsius to Kelvin offset *)
    DL_RGAS    : REAL := 8.314;    (* 通用气体常数 [J/(mol·K)] Universal gas constant *)
    DL_EXP_MAX : REAL := 50.0;     (* 指数项上钳位 [-] Exponent upper clamp *)
    DL_EXP_MIN : REAL := -50.0;    (* 指数项下钳位 [-] Exponent lower clamp *)
END_VAR
VAR
    fTK     : REAL;   (* 绝对温度 [K] Absolute temperature *)
    fTRefK  : REAL;   (* 参考绝对温度 [K] Reference absolute temperature *)
    fExp    : REAL;   (* Arrhenius 指数项 [-] Arrhenius exponent *)
END_VAR
(* 出口预置：四出口统一预置 *)
fCaseMm := 0.0; fKCoef := 0.0; fTimeTargetH := 0.0; xValid := FALSE;
(* 非有限拦截：自反判 NaN，自身差值判 Inf *)
IF (fTempC <> fTempC) OR ((fTempC - fTempC) <> 0.0)
   OR (fHoldH <> fHoldH) OR ((fHoldH - fHoldH) <> 0.0)
   OR (fKRefMmSqh <> fKRefMmSqh) OR ((fKRefMmSqh - fKRefMmSqh) <> 0.0)
   OR (fEnergyJmol <> fEnergyJmol) OR ((fEnergyJmol - fEnergyJmol) <> 0.0)
   OR (fTRefC <> fTRefC) OR ((fTRefC - fTRefC) <> 0.0)
   OR (fTargetMm <> fTargetMm) OR ((fTargetMm - fTargetMm) <> 0.0) THEN
    FC_DL_CarburizeCaseDepthCalc := -1.0;   (* 哨兵 -1：输入非有限 / Sentinel -1 non-finite *)
    RETURN;
END_IF
(* 组态域闸：保温时长非负、参考系数正、激活能非负、反算温度可表 *)
fTK := fTempC + DL_KELVIN;
fTRefK := fTRefC + DL_KELVIN;
IF (fHoldH < 0.0) OR (fKRefMmSqh <= DL_EPS) OR (fEnergyJmol < 0.0)
   OR (fTK <= DL_EPS) OR (fTRefK <= DL_EPS) THEN
    FC_DL_CarburizeCaseDepthCalc := -1.0;   (* 哨兵 -1：组态非法 / Sentinel -1 bad config *)
    RETURN;
END_IF
(* Arrhenius 温度修正：K = Kref * exp(-(Q/R)*(1/T - 1/Tref)) *)
fExp := -(fEnergyJmol / DL_RGAS) * ((1.0 / fTK) - (1.0 / fTRefK));
IF fExp > DL_EXP_MAX THEN
    fExp := DL_EXP_MAX;                     (* 指数上钳位，防 EXP 上溢 [-] / Clamp high *)
ELSIF fExp < DL_EXP_MIN THEN
    fExp := DL_EXP_MIN;                     (* 指数下钳位，防 EXP 下溢 [-] / Clamp low *)
END_IF
fKCoef := fKRefMmSqh * EXP(fExp);           (* 当前温度 K 系数 [mm/sqrt(h)] / K at temperature *)
(* Harris 层深：x = K*sqrt(t)，开方前已保证 t >= 0 *)
fCaseMm := fKCoef * SQRT(fHoldH);
(* 反算保温时间：t = (x/K)^2，K 已过域闸 *)
IF fTargetMm > 0.0 THEN
    fTimeTargetH := (fTargetMm / fKCoef) * (fTargetMm / fKCoef);
END_IF
(* 输出自检：K 极小或 t 极大时 (x/K)^2 可上溢 Inf，出口一律复检非有限 *)
IF (fCaseMm <> fCaseMm) OR ((fCaseMm - fCaseMm) <> 0.0)
   OR (fKCoef <= DL_EPS)
   OR (fTimeTargetH <> fTimeTargetH) OR ((fTimeTargetH - fTimeTargetH) <> 0.0) THEN
    fCaseMm := 0.0; fKCoef := 0.0; fTimeTargetH := 0.0;
    xValid := FALSE;                         (* 输出不可信 / Output not trustworthy *)
    FC_DL_CarburizeCaseDepthCalc := -1.0;    (* 哨兵 -1：输出溢出 / Sentinel -1 overflow *)
    RETURN;
END_IF
xValid := TRUE;                             (* 链路有效 / Chain valid *)
FC_DL_CarburizeCaseDepthCalc := fCaseMm;    (* 返回层深 [mm] / Return case depth *)
END_FUNCTION

(* ---- FC_DL_CasingRateCalc.st ---- *)
(*
 * FC_DL_CasingRateCalc | C2 | DL_Process
 * 功能：叶片加料比例与实际料液体积流量（按料液密度换算）       单位：流量 [kg/h]、比例 [%]、密度 [kg/L]、体积流量 [L/h]
 * 工况边界：叶片流量须 >0（入分母）；料液密度取 1.05 kg/L 固定常数（糖香料液典型值），密度差异超出 ±0.05 须现场标定；料液流量不得为负
 * 代数值回代：leaf=5000 kg/h、casing=150 kg/h → rate=150/5000×100=3.0 %（=目标 3.0 %，合格）；flow=150/1.05=142.9 L/h（与 spec 比例式一致）
 * 开源溯源：clean-room 自研，未复制任何第三方代码（无外部来源）
 *)
FUNCTION FC_DL_CasingRateCalc : BOOL
VAR_INPUT
    rLeafKgH     : REAL := 5000.0;   // 叶片流量 | leaf tobacco mass flow [kg/h]
    rCasingKgH   : REAL;             // 料液质量流量 | casing mass flow [kg/h]
    rTargetPct   : REAL := 3.0;      // 目标加料比例 | target casing ratio [%]
    rTolPct      : REAL := 0.2;      // 加料比例公差（±）| casing ratio tolerance [%]
END_VAR
VAR_OUTPUT
    rRatePct      : REAL;            // 实际加料比例 | actual casing ratio [%]
    rCasingFlowLh : REAL;            // 料液体积流量（按密度换算）| casing volumetric flow [L/h]
    rDevPct       : REAL;            // 相对目标的偏差 | deviation from the target [%]
    xInTolerance  : BOOL;            // 比例在公差带内 | ratio within tolerance
    xValid        : BOOL;            // 输出有效 | outputs valid
END_VAR
VAR
    xFinLeaf : BOOL;                 // 叶片流量有限性 | leaf flow is finite
    xFinCase : BOOL;                 // 料液流量有限性 | casing flow is finite
    xFinTg   : BOOL;                 // 目标有限性 | target is finite
    xFinTol  : BOOL;                 // 公差有限性 | tolerance is finite
END_VAR
VAR CONSTANT
    DL_CRC_PCT   : REAL := 100.0;    // 百分数换算系数 | percentage factor [%]
    DL_CRC_DENS  : REAL := 1.05;     // 料液密度（固定常数，需现场标定）| casing density, a fixed constant to be calibrated on site [kg/L]
    DL_CRC_DMIN  : REAL := 1.0E-9;   // 除零保护阈值 | division guard threshold [kg/h]
    DL_CRC_EPS   : REAL := 1.0E-6;   // 浮点比较容差 | floating comparison tolerance [%]
END_VAR

// 段1｜非有限闸（R19）
xFinLeaf := (rLeafKgH = rLeafKgH) AND ((rLeafKgH - rLeafKgH) = 0.0);
xFinCase := (rCasingKgH = rCasingKgH) AND ((rCasingKgH - rCasingKgH) = 0.0);
xFinTg := (rTargetPct = rTargetPct) AND ((rTargetPct - rTargetPct) = 0.0);
xFinTol := (rTolPct = rTolPct) AND ((rTolPct - rTolPct) = 0.0);
IF (NOT xFinLeaf) OR (NOT xFinCase) OR (NOT xFinTg) OR (NOT xFinTol) THEN
    rRatePct := 0.0;                 // 安全值：比例 0 | safe value, zero ratio
    rCasingFlowLh := 0.0;
    rDevPct := 0.0;
    xInTolerance := FALSE;
    xValid := FALSE;
    FC_DL_CasingRateCalc := FALSE;
    RETURN;
END_IF

// 段2｜域闸：叶片流量 >0、料液流量 ≥0、公差 ≥0
IF (rLeafKgH <= DL_CRC_DMIN) OR (rCasingKgH < 0.0) OR (rTolPct < 0.0) THEN
    rRatePct := 0.0;
    rCasingFlowLh := 0.0;
    rDevPct := 0.0;
    xInTolerance := FALSE;
    xValid := FALSE;
    FC_DL_CasingRateCalc := FALSE;
    RETURN;
END_IF

// 段3｜算法：rate = casing/leaf×100；体积流量 = 质量流量/密度
rRatePct := rCasingKgH / rLeafKgH * DL_CRC_PCT;
rCasingFlowLh := rCasingKgH / DL_CRC_DENS;     // 密度为常数 1.05，恒非零 | the density constant is never zero

// 段4｜合格判定（判据与出口同源于原始流量）
rDevPct := rRatePct - rTargetPct;
xInTolerance := ABS(rDevPct) <= (rTolPct + DL_CRC_EPS);
xValid := TRUE;
FC_DL_CasingRateCalc := TRUE;
END_FUNCTION

(* ---- FC_DL_CastingSolidificationTimeCalc.st ---- *)
(*
  Component : FC_DL_CastingSolidificationTimeCalc
  Category  : DL_Process
  Type      : FC
  Complexity: C1
  VERSION   : v1.0.0
  功能      : Chvorinov 凝固时间核算：t = B·(V/A)² 算铸件凝固时间，并由铸件模数与冷铁判据判断是否需要加冷铁。
  开源溯源  : 道莅原创 clean-room 自研（无外部代码引用）｜License: MIT
  边界条件  : ① 铸件体积与散热表面积须 > 1e-9，否则返回哨兵 -1（体积按 cm³、面积按 cm² 输入）；
              ② 冷铁判据以模数为唯一依据：模数大于临界模数即建议加冷铁；
              ③ 凝固时间常数 B 须为正，负值判组态非法。
*)
FUNCTION FC_DL_CastingSolidificationTimeCalc : REAL
VAR_INPUT
    fVolCm3        : REAL;   (* 铸件体积 [cm³] Casting volume *)
    fSurfAreaCm2   : REAL;   (* 有效散热表面积 [cm²] Effective cooling surface *)
    fChvorinovBS   : REAL;   (* Chvorinov 时间常数 [s/cm²] Chvorinov constant *)
    fModulusCritCm : REAL;   (* 冷铁判据临界模数 [cm] Critical modulus for chill *)
END_VAR
VAR_OUTPUT
    fModulusCm  : REAL;   (* 铸件模数 V/A [cm] Casting modulus *)
    fSolidTimeS : REAL;   (* 凝固时间 [s] Solidification time *)
    xNeedChill  : BOOL;   (* 建议加冷铁标志 [-] Chill recommended flag *)
    xValid      : BOOL;   (* 计算有效性标志 [-] Calculation valid flag *)
END_VAR
VAR CONSTANT
    DL_EPS  : REAL := 1.0E-9;   (* 除零判定容差 [无量纲] Divide-by-zero tolerance *)
    DL_ZERO : REAL := 0.0;      (* 零常量 [无量纲] Zero constant *)
END_VAR
(* 出口预置：四出口统一预置 *)
fModulusCm := 0.0; fSolidTimeS := 0.0; xNeedChill := FALSE; xValid := FALSE;
(* 非有限拦截：自反判 NaN，自身差值判 Inf *)
IF (fVolCm3 <> fVolCm3) OR ((fVolCm3 - fVolCm3) <> 0.0)
   OR (fSurfAreaCm2 <> fSurfAreaCm2) OR ((fSurfAreaCm2 - fSurfAreaCm2) <> 0.0)
   OR (fChvorinovBS <> fChvorinovBS) OR ((fChvorinovBS - fChvorinovBS) <> 0.0)
   OR (fModulusCritCm <> fModulusCritCm) OR ((fModulusCritCm - fModulusCritCm) <> 0.0) THEN
    FC_DL_CastingSolidificationTimeCalc := -1.0;  (* 哨兵 -1：输入非有限 / Sentinel -1 non-finite *)
    RETURN;
END_IF
(* 组态域闸：体积、面积均为除子或比例基，时间常数须为正 *)
IF (fVolCm3 <= DL_EPS) OR (fSurfAreaCm2 <= DL_EPS) OR (fChvorinovBS <= DL_ZERO)
   OR (fModulusCritCm <= DL_ZERO) THEN
    FC_DL_CastingSolidificationTimeCalc := -1.0;  (* 哨兵 -1：组态非法 / Sentinel -1 bad config *)
    RETURN;
END_IF
(* 铸件模数：M = V/A [cm]，分母已过域闸 *)
fModulusCm := fVolCm3 / fSurfAreaCm2;
(* Chvorinov：t = B·M² [s] *)
fSolidTimeS := fChvorinovBS * fModulusCm * fModulusCm;
(* 冷铁判据：模数超过临界模数即建议局部加冷铁 *)
xNeedChill := fModulusCm > fModulusCritCm;
xValid := TRUE;                                 (* 链路有效 / Chain valid *)
FC_DL_CastingSolidificationTimeCalc := fSolidTimeS;  (* 返回凝固时间 [s] / Return solidification time *)
END_FUNCTION

(* ---- FC_DL_CatalystActivityDecay.st ---- *)
(*
  道莅工业代码库 / Daoli Industrial ST Library
  组件: FC_DL_CatalystActivityDecay
  分类: DL_Process
  开源溯源: 无（clean-room 工程公式自研；参考公开工艺计算公式，未复制任何受版权保护代码）
  许可证: 本项目自有 (MIT)
  功能: 催化剂活性一阶衰减模型：活性、温度加速失活因子与剩余可用寿命 RUL
  模型: k = k0·EXP(Kt·(T-Tref))；act = EXP(-k·t)；RUL = (k·t + LN(1/0.7))/k
*)
FUNCTION FC_DL_CatalystActivityDecay : BOOL
VAR_INPUT
    rDeactBase : REAL; // 基准温度下失活速率常数 [1/h] / base deactivation rate constant
    rHoursRun : REAL; // 累计运行小时数 [h] / accumulated operating hours
    rTempC : REAL; // 实际运行温度 [°C] / actual operating temperature
    rTempRefC : REAL; // 基准温度 [°C] / reference temperature
    rKt : REAL; // 温度加速系数 [1/°C] / temperature acceleration coefficient
END_VAR
VAR_OUTPUT
    rActivity : REAL; // 相对活性 [-]，1.0 = 全新 / relative activity, 1.0 is fresh
    rRulHours : REAL; // 活性降至 0.7 的剩余小时数 [h] / remaining useful life to 70 percent activity
    bValid : BOOL; // 结果有效位 [-] / result valid flag
    iErrCode : INT; // 事件码 0=正常 1=基准失活率非法 2=失活率近零无退化 3=运行小时为负 4=温度低于绝对零度 5=结果非有限 / event code
END_VAR
VAR CONSTANT
    rLnInv07 : REAL := 0.356674944; // LN(1/0.7) 寿命终点常数 [-] / LN of one over 0.7
    rActFloor : REAL := 0.0001; // 活性下限 [-]，防 LN(0) / activity floor preventing LN of zero
    rActCeil : REAL := 1.0; // 活性上限 [-]，不得高于全新 / activity ceiling, never above fresh
    rExpHi : REAL := 50.0; // EXP 指数量程上限 [-]，防溢出 / exponent ceiling guarding EXP overflow
    rExpLo : REAL := -50.0; // EXP 指数量程下限 [-] / exponent floor
    rKelvinOff : REAL := 273.15; // 开尔文偏移 [K] / kelvin offset
END_VAR
VAR
    rExpo : REAL; // 温度加速指数 [-] / temperature exponent
    rK : REAL; // 实际失活速率常数 [1/h] / effective deactivation rate constant
    rAct : REAL; // 未限幅活性 [-] / unlimited activity
    rRulRaw : REAL; // 未限幅剩余寿命 [h] / unlimited remaining life
END_VAR

    // —— 段 0：全路径预清 —— //
    rExpo := 0.0;
    rK := 0.0;
    rAct := 0.0;
    rRulRaw := 0.0;
    rActivity := rActFloor;
    rRulHours := 0.0;
    bValid := FALSE;
    iErrCode := 0;
    FC_DL_CatalystActivityDecay := FALSE;
    // —— 段 1：输入域闸 —— //
    IF rDeactBase <= 0.0 THEN
        iErrCode := 1; // 基准失活率非法，衰减模型无定义 / invalid base rate, model undefined
        RETURN;
    END_IF;
    IF rHoursRun < 0.0 THEN
        iErrCode := 3; // 运行小时为负 / negative operating hours
        RETURN;
    END_IF;
    IF rTempC <= (0.0 - rKelvinOff) THEN
        iErrCode := 4; // 温度低于绝对零度，物理不可能 / temperature below absolute zero
        RETURN;
    END_IF;
    // —— 段 2：温度加速失活常数（指数先做量程钳位，防 EXP 溢出） —— //
    rExpo := rKt * (rTempC - rTempRefC); // 加速指数 [-] / acceleration exponent
    IF rExpo > rExpHi THEN
        rExpo := rExpHi; // 上限钳位 / clamp high
    ELSIF rExpo < rExpLo THEN
        rExpo := rExpLo; // 下限钳位 / clamp low
    END_IF;
    rK := rDeactBase * EXP(rExpo); // 失活速率常数 [1/h] / rate constant
    // —— 段 3：活性 = EXP(-k·t)，并限 [0.0001, 1] —— //
    rAct := EXP(0.0 - rK * rHoursRun); // 活性 [-] / activity
    IF rAct > rActCeil THEN
        rActivity := rActCeil; // 上限钳位 / clamp high
    ELSIF rAct < rActFloor THEN
        rActivity := rActFloor; // 下限钳位，保证后续 LN 有定义 / floor keeps LN defined
    ELSE
        rActivity := rAct;
    END_IF;
    // —— 段 4：RUL（分母闸：k 必须显著为正；LN 前闸：活性为正） —— //
    IF rK <= 1.0E-9 THEN
        rRulHours := 99999.0; // 失活率近零，视为无退化 / near-zero decay, treat as no degradation
        iErrCode := 2; // 信息级：无退化，寿命取哨兵值 / info: no degradation, sentinel life
        bValid := TRUE;
        FC_DL_CatalystActivityDecay := TRUE;
        RETURN;
    END_IF;
    IF rActivity <= 0.0 THEN
        iErrCode := 5; // 活性非正，LN 无定义 / non-positive activity, LN undefined
        RETURN;
    END_IF;
    // 量纲 (-)/(1/h) = h；目标时刻 LN(1/0.7)/k 减去已运行量 LN(1/act)/k
    rRulRaw := (rLnInv07 - LN(1.0 / rActivity)) / rK; // 剩余寿命 [h] / remaining life in hours
    IF ABS(rRulRaw) > 1.0E15 THEN
        rRulHours := 0.0;
        iErrCode := 5; // 结果非有限，强制归零 / non-finite result, forced to zero
        RETURN;
    END_IF;
    IF rRulRaw < 0.0 THEN
        rRulHours := 0.0; // 已过寿命终点 / life already exhausted
    ELSE
        rRulHours := rRulRaw;
    END_IF;
    bValid := TRUE;
    FC_DL_CatalystActivityDecay := TRUE;
END_FUNCTION

(* ---- FC_DL_CathodeD50TargetCalc.st ---- *)
(*
  Component : FC_DL_CathodeD50TargetCalc
  Category  : DL_Process
  Function  : 目标 D50 与分级轮转速反算：d50 = k / rpm，含上下限钳位
  Complexity: C2
  开源溯源 : DLF 内部原创（R94 族模板派生）；参考语义来源见 SOURCE_HUNTING_MATRIX.md
  规则遵从 : R1-R16
  契约     : 输入 nWheelRpm 分级轮转速 [r/min]、rCoefUmRpm 切割系数 [μm·r/min]、
             rD50MinUm 目标下限 [μm]、rD50MaxUm 目标上限 [μm]；
             输出 rD50Um 钳位后目标 D50 [μm]、rD50RawUm 未钳位计算值 [μm]、
             xClamped 触限、xValid 有效标志、nFaultCode 故障码。
  边界     : 转速为分母须 >1（转速过低无切割效应，模型外推发散）；上下限须 上限 > 下限 > 0；
             切割系数须 >1.0E-9 [μm·r/min]；钳位后仍给出未钳位值以便上层判断模型是否越界。
  码位     : 9801 输入非有限（故障级）；9802 转速、系数或限值越域（故障级）。
*)
FUNCTION FC_DL_CathodeD50TargetCalc : BOOL
VAR_INPUT
    nWheelRpm  : INT := 3000;        // 分级轮转速 [r/min] EN: the rotational speed of the classifying wheel
    rCoefUmRpm : LREAL := 30000.0;   // 切割系数（D50 × 转速） [μm·r/min] EN: the cut coefficient, the product of D50 and the speed
    rD50MinUm  : LREAL := 1.0;       // 目标 D50 下限 [μm] EN: the lower bound of the target median size
    rD50MaxUm  : LREAL := 30.0;      // 目标 D50 上限 [μm] EN: the upper bound of the target median size
END_VAR
VAR_OUTPUT
    rD50Um    : LREAL;               // 钳位后目标 D50 [μm] EN: the clamped target median size
    rD50RawUm : LREAL;               // 未钳位计算值 [μm] EN: the unclamped computed median size
    xClamped  : BOOL;                // 触上下限 EN: the bound was reached
    xValid    : BOOL;                // 输出可信标志 EN: the outputs are valid
    nFaultCode: INT;                 // 0=无故障 9801=输入非有限 9802=转速或限值越域 EN: zero none, 9801 non finite, 9802 speed or limits out of range
END_VAR
VAR
    xFinAll : BOOL;                  // 浮点入参有限 EN: the floating inputs are finite
    rDen    : LREAL;                 // 分母（转速实数化） [r/min] EN: the divisor, the speed as a real number
    rRaw    : LREAL;                 // 计算中间值 [μm] EN: the interim computed value
    rOut    : LREAL;                 // 钳位后中间值 [μm] EN: the interim clamped value
END_VAR
VAR CONSTANT
    DL_CDT_Z     : LREAL := 0.0;     // 浮点零常量 EN: the floating point zero constant
    DL_CDT_ONE   : LREAL := 1.0;     // 浮点壹常量 EN: the floating point one constant
    DL_CDT_MIN   : LREAL := 1.0E-9;  // 分母绝对值下限 EN: the lower bound of the divisor magnitude
    DL_CDT_C_BAD : INT := 9801;      // 输入非有限 EN: a non finite input
    DL_CDT_C_RANG: INT := 9802;      // 转速或限值越域 EN: the speed or the limits are out of range
END_VAR

// 段1｜出口预置
FC_DL_CathodeD50TargetCalc := FALSE;   // 返回值预置假 EN: preset the return value to false
rD50Um := DL_CDT_Z;                    // 钳位值预置零 [μm] EN: preset the clamped value to zero
rD50RawUm := DL_CDT_Z;                 // 未钳位值预置零 [μm] EN: preset the unclamped value to zero
xClamped := FALSE;                     // 触限标志预置假 EN: preset the clamp flag to false
xValid := FALSE;                       // 有效标志预置假 EN: preset the validity flag to false
nFaultCode := 0;                       // 故障码预置零 EN: preset the fault code to zero

// 段2｜非有限闸：三浮点入参全列（两限值参与钳位）
xFinAll := (rCoefUmRpm = rCoefUmRpm) AND ((rCoefUmRpm - rCoefUmRpm) = DL_CDT_Z)
        AND (rD50MinUm = rD50MinUm) AND ((rD50MinUm - rD50MinUm) = DL_CDT_Z)
        AND (rD50MaxUm = rD50MaxUm) AND ((rD50MaxUm - rD50MaxUm) = DL_CDT_Z);   // 三输入有限性 EN: the finiteness of all three inputs
IF NOT xFinAll THEN                                                             // 非有限出口 EN: leave early on a non finite input
    nFaultCode := DL_CDT_C_BAD;                                                 // 非有限码 EN: the non finite code
    RETURN;                                                                     // 早退 EN: return early
END_IF

// 段3｜域闸：转速 >1 [r/min]、系数为正、限值 上限 > 下限 > 0
rDen := INT_TO_LREAL(nWheelRpm);                                                // 转速实数化 [r/min] EN: the speed as a real number
IF (rDen <= DL_CDT_ONE) OR (ABS(rCoefUmRpm) < DL_CDT_MIN)
   OR (rD50MinUm <= DL_CDT_Z) OR (rD50MaxUm <= rD50MinUm) THEN
    nFaultCode := DL_CDT_C_RANG;                                                // 越域码 EN: the out of range code
    RETURN;                                                                     // 早退 EN: return early
END_IF

// 段4｜主体：d50 = k / rpm
rRaw := rCoefUmRpm / rDen;                                                      // 计算 D50 [μm] EN: the computed median size
IF (rRaw <> rRaw) OR (rRaw <= DL_CDT_Z) THEN                                    // 结果复检 EN: recheck the result
    nFaultCode := DL_CDT_C_RANG;                                                // 复检失败码 EN: the recheck failure code
    RETURN;                                                                     // 早退，出口保持零哨兵 EN: return early with the zero sentinels
END_IF

// 段5｜上下限钳位（不饱和报表：xClamped 表达模型是否越界）
rOut := rRaw;                                                                   // 钳位工作副本 [μm] EN: the working copy for clamping
IF rOut < rD50MinUm THEN                                                        // 下钳位 EN: clamp the lower bound
    rOut := rD50MinUm;                                                          // 抬到下限 [μm] EN: raise to the lower bound
    xClamped := TRUE;                                                           // 置触限标志 EN: raise the clamp flag
END_IF
IF rOut > rD50MaxUm THEN                                                        // 上钳位 EN: clamp the upper bound
    rOut := rD50MaxUm;                                                          // 压到上限 [μm] EN: clamp to the upper bound
    xClamped := TRUE;                                                           // 置触限标志 EN: raise the clamp flag
END_IF

// 段6｜出口
rD50Um := rOut;                                                                 // 钳位值出口 [μm] EN: the clamped value output
rD50RawUm := rRaw;                                                              // 未钳位值出口 [μm] EN: the unclamped value output
xValid := TRUE;                                                                 // 结果可信 EN: the results are valid
FC_DL_CathodeD50TargetCalc := TRUE;                                             // 返回真 EN: return true
END_FUNCTION

(* ---- FC_DL_CathodeLiExcessCalc.st ---- *)
(*
  Component : FC_DL_CathodeLiExcessCalc
  Category  : DL_Process
  Function  : 锂电正极材料 Li/M 摩尔比与实际过量率，并做目标区间判定
  Complexity: C2
  开源溯源 : DLF 内部原创（R94 族模板派生）；参考语义来源见 SOURCE_HUNTING_MATRIX.md
  规则遵从 : R1-R16
  契约     : 输入 rLiMolPerM 实测 Li/M 摩尔比 [-]、rTargetRatio 目标 Li/M 摩尔比 [-]、
             rBandTolPct 目标区间半宽 [%]；输出 rExcessPct 相对目标过量率 [%]、rLiMolPerM 摩尔比直通、
             xInBand 摩尔比落在目标区间、xValid 有效标志、nFaultCode 故障码。
  边界     : 目标摩尔比为分母须 >1.0E-9；区间半宽须在 (0, 50] [%] 内，越域判 9803（半宽越域使判定
             恒真或恒假，属组态域闸缺失）；过量率可正可负，负值表达欠锂，不做钳位（方向信息不得丢失）。
  码位     : 9801 输入非法（故障级）；9802 目标摩尔比过小（故障级）；9803 区间半宽越域（故障级）。
*)
FUNCTION FC_DL_CathodeLiExcessCalc : BOOL
VAR_INPUT
    rLiMolPerM    : LREAL := 1.03;   // 实测 Li/M 摩尔比 [-] EN: the measured lithium to metal molar ratio
    rTargetRatio  : LREAL := 1.03;   // 目标 Li/M 摩尔比 [-] EN: the target lithium to metal molar ratio
    rBandTolPct   : LREAL := 1.0;    // 目标区间半宽 [%] EN: the half width of the target band in percent
END_VAR
VAR_OUTPUT
    rExcessPct  : LREAL;             // 相对目标摩尔比的过量率 [%] EN: the excess rate against the target molar ratio
    rRatioEcho  : LREAL;             // 摩尔比直通（供趋势记录） [-] EN: the molar ratio passed through for trending
    xInBand     : BOOL;              // 摩尔比落在目标区间 EN: the molar ratio is inside the target band
    xValid      : BOOL;              // 输出可信标志 EN: the outputs are valid
    nFaultCode  : INT;               // 0=无故障 9801=输入非法 9802=目标比过小 9803=半宽越域 EN: zero none, 9801 illegal input, 9802 target too small, 9803 half width out of range
END_VAR
VAR
    xFinAll  : BOOL;                 // 三输入同时有限 EN: all three inputs are finite
    rDev     : LREAL;                // 相对偏差 [-] EN: the relative deviation
    rDevPct  : LREAL;                // 相对偏差百分数 [%] EN: the relative deviation in percent
    rDen     : LREAL;                // 分母（目标摩尔比） [-] EN: the divisor, the target molar ratio
END_VAR
VAR CONSTANT
    DL_CLE_Z       : LREAL := 0.0;   // 浮点零常量 EN: the floating point zero constant
    DL_CLE_HUNDRED : LREAL := 100.0; // 百分数换算系数 EN: the percent conversion factor
    DL_CLE_TOL_MAX : LREAL := 50.0;  // 区间半宽上限 [%] EN: the upper bound of the band half width
    DL_CLE_MIN     : LREAL := 1.0E-9;// 分母绝对值下限 EN: the lower bound of the divisor magnitude
    DL_CLE_C_BAD   : INT := 9801;    // 输入非法 EN: an illegal input
    DL_CLE_C_TGT   : INT := 9802;    // 目标摩尔比过小 EN: the target molar ratio is too small
    DL_CLE_C_TOL   : INT := 9803;    // 区间半宽越域 EN: the half width is out of range
END_VAR

// 段1｜出口预置
FC_DL_CathodeLiExcessCalc := FALSE;   // 返回值预置假 EN: preset the return value to false
rExcessPct := DL_CLE_Z;                // 过量率预置零 [%] EN: preset the excess rate to zero
rRatioEcho := DL_CLE_Z;                // 摩尔比直通预置零 [-] EN: preset the ratio echo to zero
xInBand := FALSE;                      // 区间标志预置假 EN: preset the band flag to false
xValid := FALSE;                       // 有效标志预置假 EN: preset the validity flag to false
nFaultCode := 0;                       // 故障码预置零 EN: preset the fault code to zero

// 段2｜非有限闸：三输入全列（半宽参与区间判据，漏则判定失效）
xFinAll := (rLiMolPerM = rLiMolPerM) AND ((rLiMolPerM - rLiMolPerM) = DL_CLE_Z)
        AND (rTargetRatio = rTargetRatio) AND ((rTargetRatio - rTargetRatio) = DL_CLE_Z)
        AND (rBandTolPct = rBandTolPct) AND ((rBandTolPct - rBandTolPct) = DL_CLE_Z);   // 三输入有限性 EN: the finiteness of all three inputs
IF NOT xFinAll THEN                                                                     // 非有限出口 EN: leave early on a non finite input
    nFaultCode := DL_CLE_C_BAD;                                                         // 输入非法码 EN: the illegal input code
    RETURN;                                                                             // 早退 EN: return early
END_IF

// 段3｜域闸：目标比为分母须过下限；半宽须在 (0,50] 内
rDen := rTargetRatio;                                                                   // 取分母 [-] EN: take the divisor
IF ABS(rDen) < DL_CLE_MIN THEN                                                          // 分母下限 EN: the divisor magnitude gate
    nFaultCode := DL_CLE_C_TGT;                                                         // 目标比过小码 EN: the target ratio code
    RETURN;                                                                             // 早退 EN: return early
END_IF
IF (rBandTolPct <= DL_CLE_Z) OR (rBandTolPct > DL_CLE_TOL_MAX) THEN                     // 半宽域闸 EN: the half width domain gate
    nFaultCode := DL_CLE_C_TOL;                                                         // 半宽越域码 EN: the half width code
    RETURN;                                                                             // 早退 EN: return early
END_IF

// 段4｜主体：过量率 = (实测/目标 − 1) × 100，不钳位以保留欠锂方向
rDev := (rLiMolPerM / rDen) - 1.0;                                                      // 相对偏差 [-] EN: the relative deviation
rDevPct := rDev * DL_CLE_HUNDRED;                                                       // 相对偏差百分数 [%] EN: the relative deviation in percent

// 段5｜出口：区间判定按绝对值比较（欠锂与过锂同带宽）
rExcessPct := rDevPct;                                                                  // 过量率出口 [%] EN: the excess rate output
rRatioEcho := rLiMolPerM;                                                               // 摩尔比直通 [-] EN: the ratio echo output
xInBand := ABS(rDevPct) <= rBandTolPct;                                                 // 区间判定 EN: the band verdict
xValid := TRUE;                                                                         // 结果可信 EN: the results are valid
FC_DL_CathodeLiExcessCalc := TRUE;                                                      // 返回真 EN: return true
END_FUNCTION
